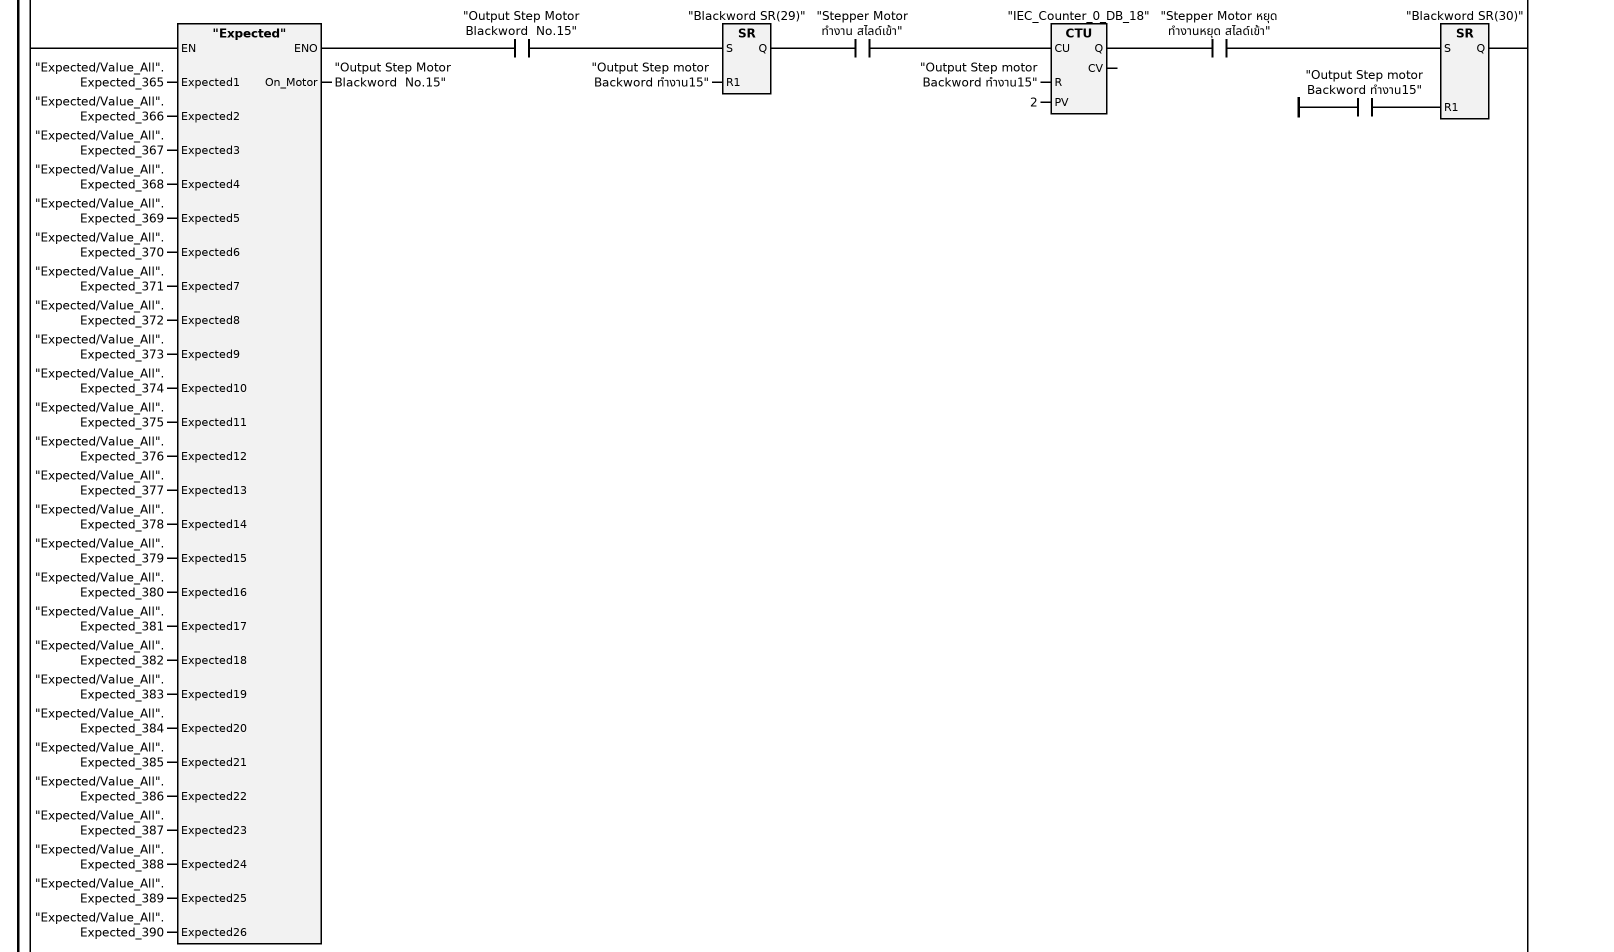
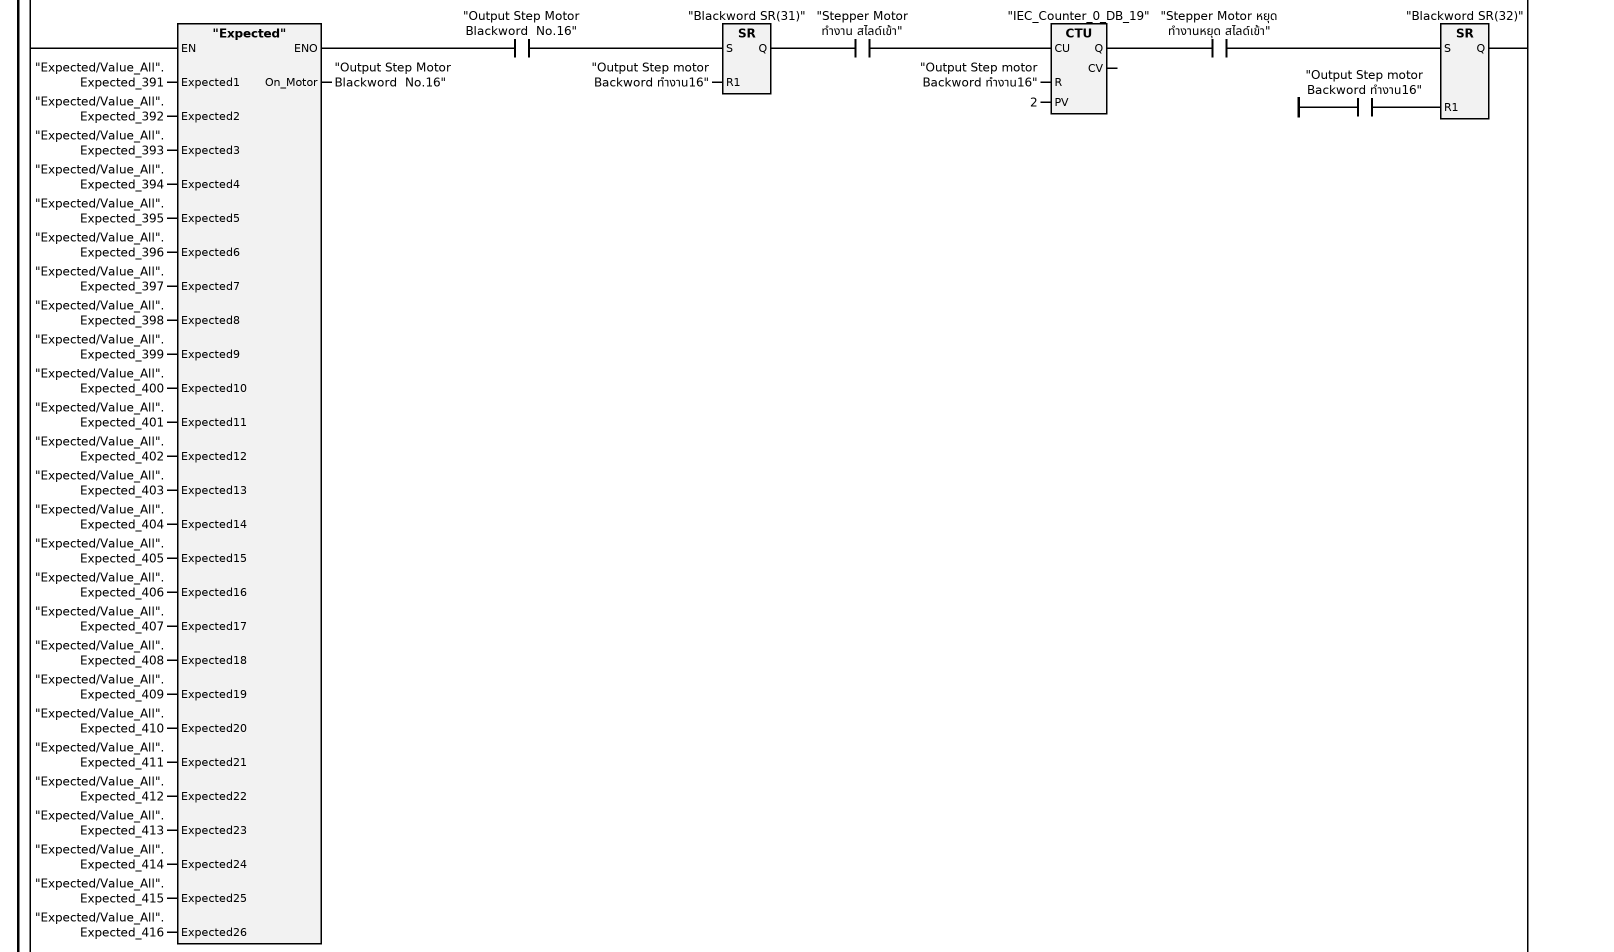
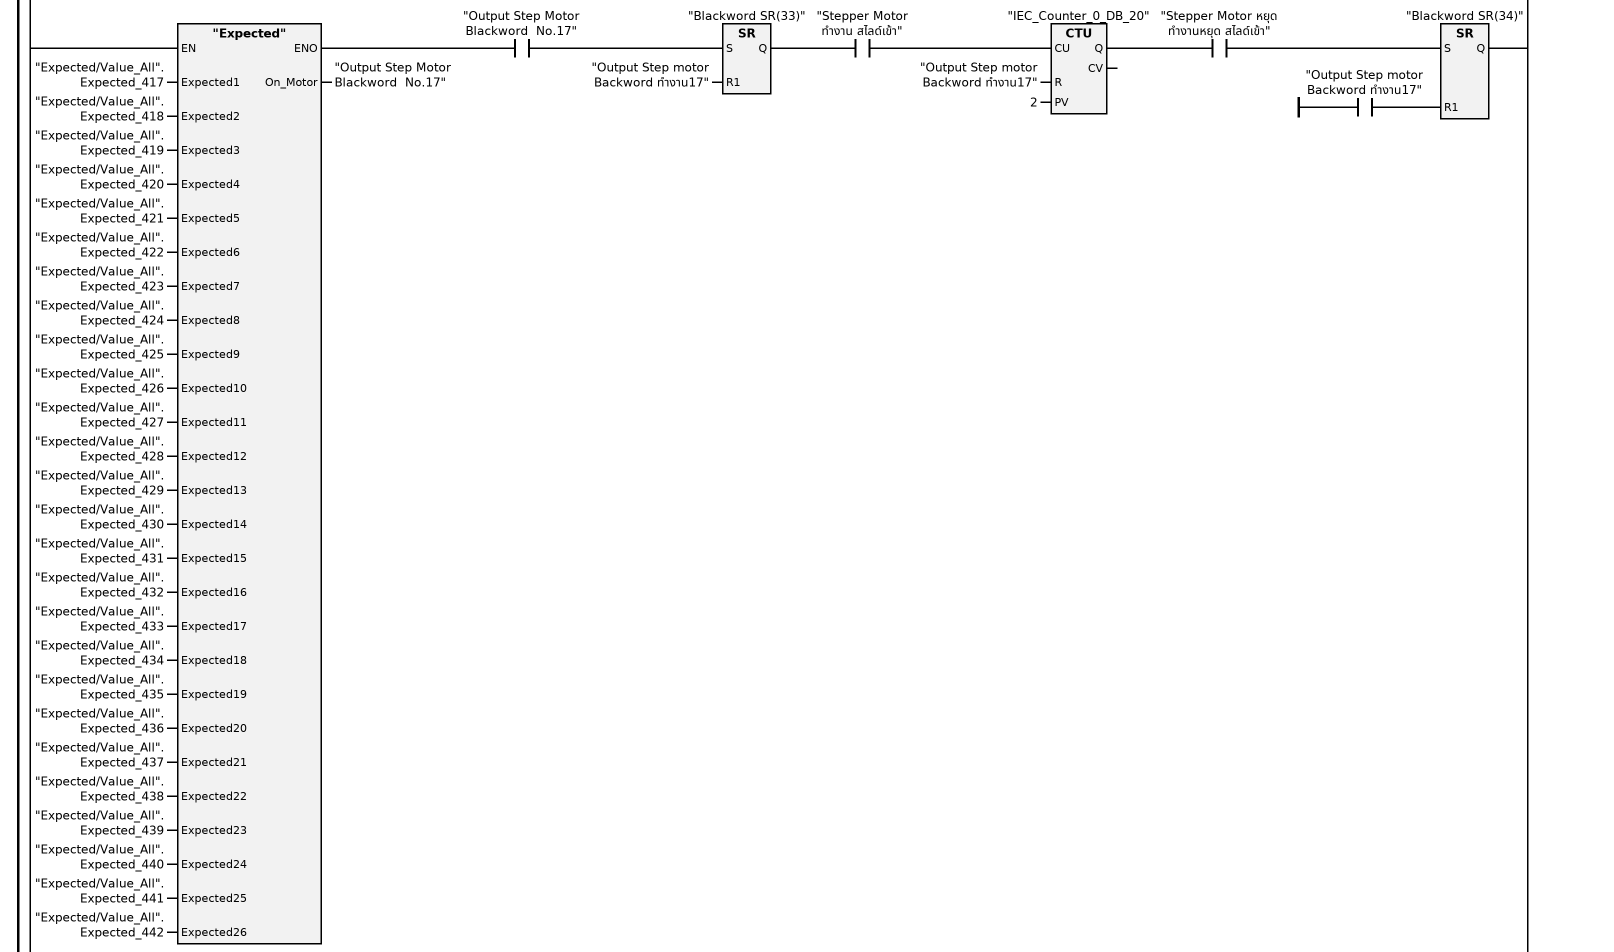
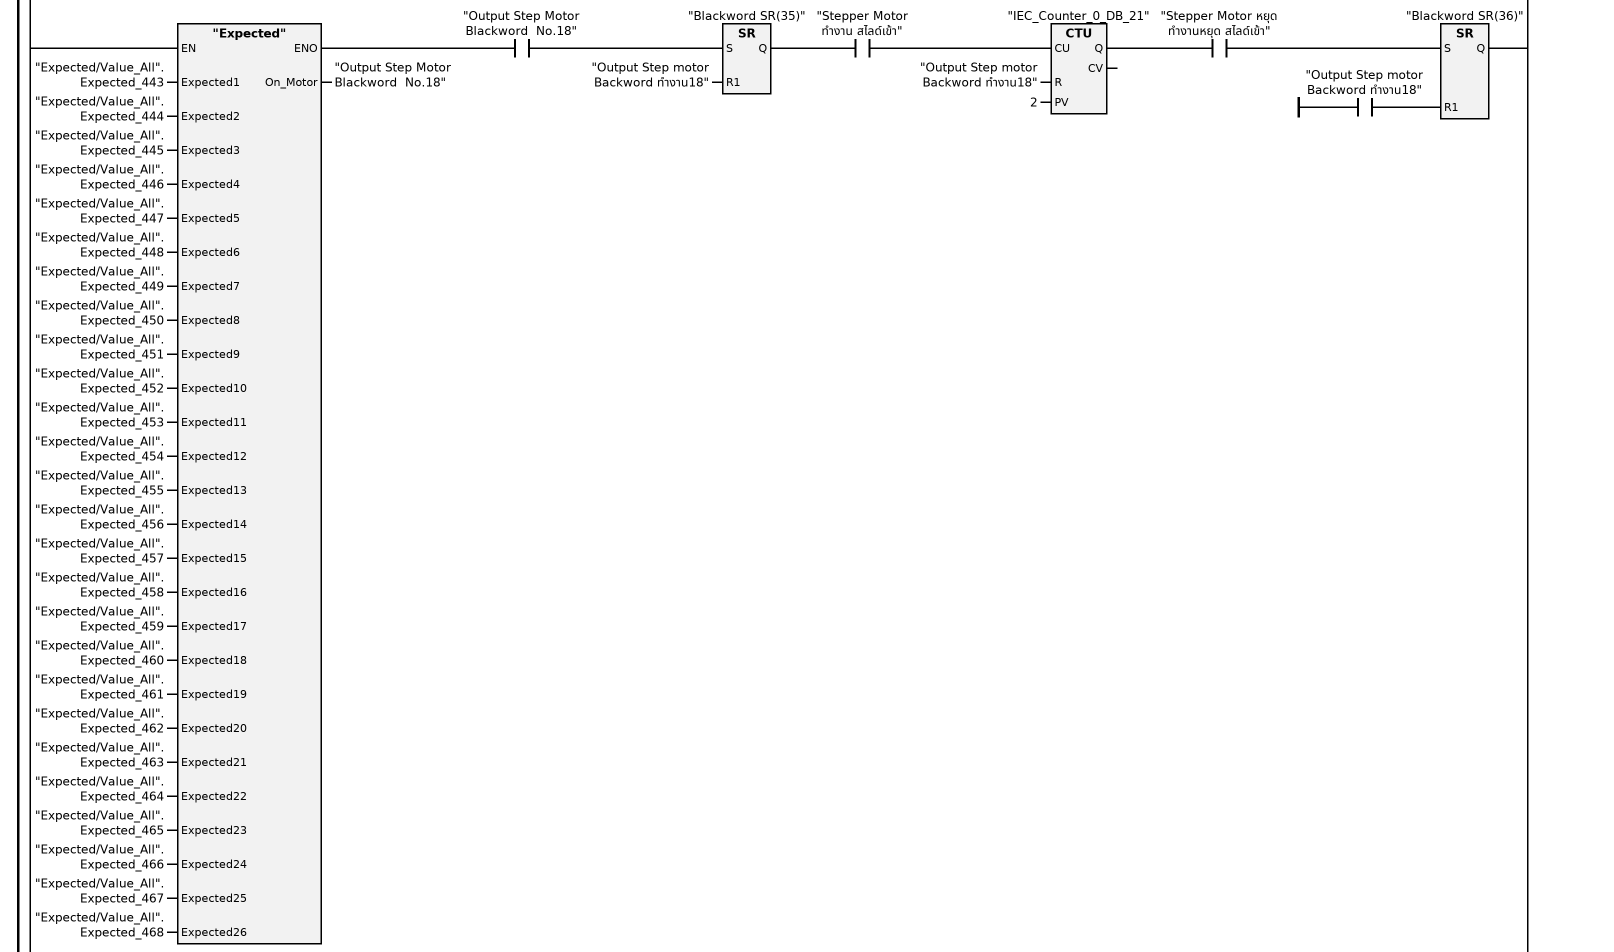
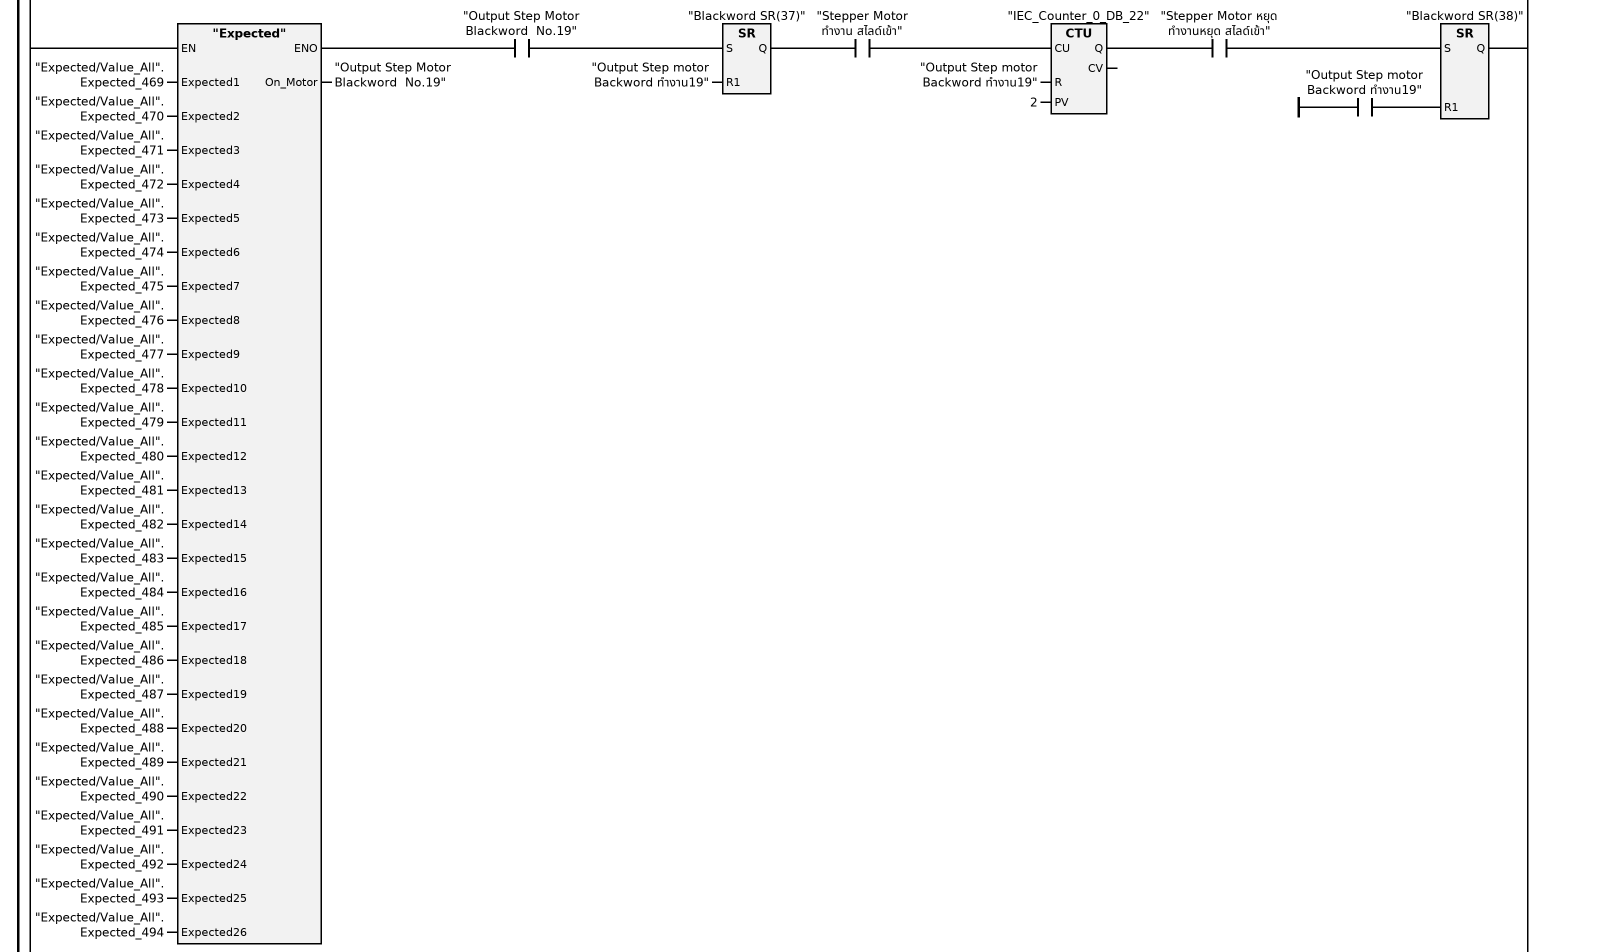
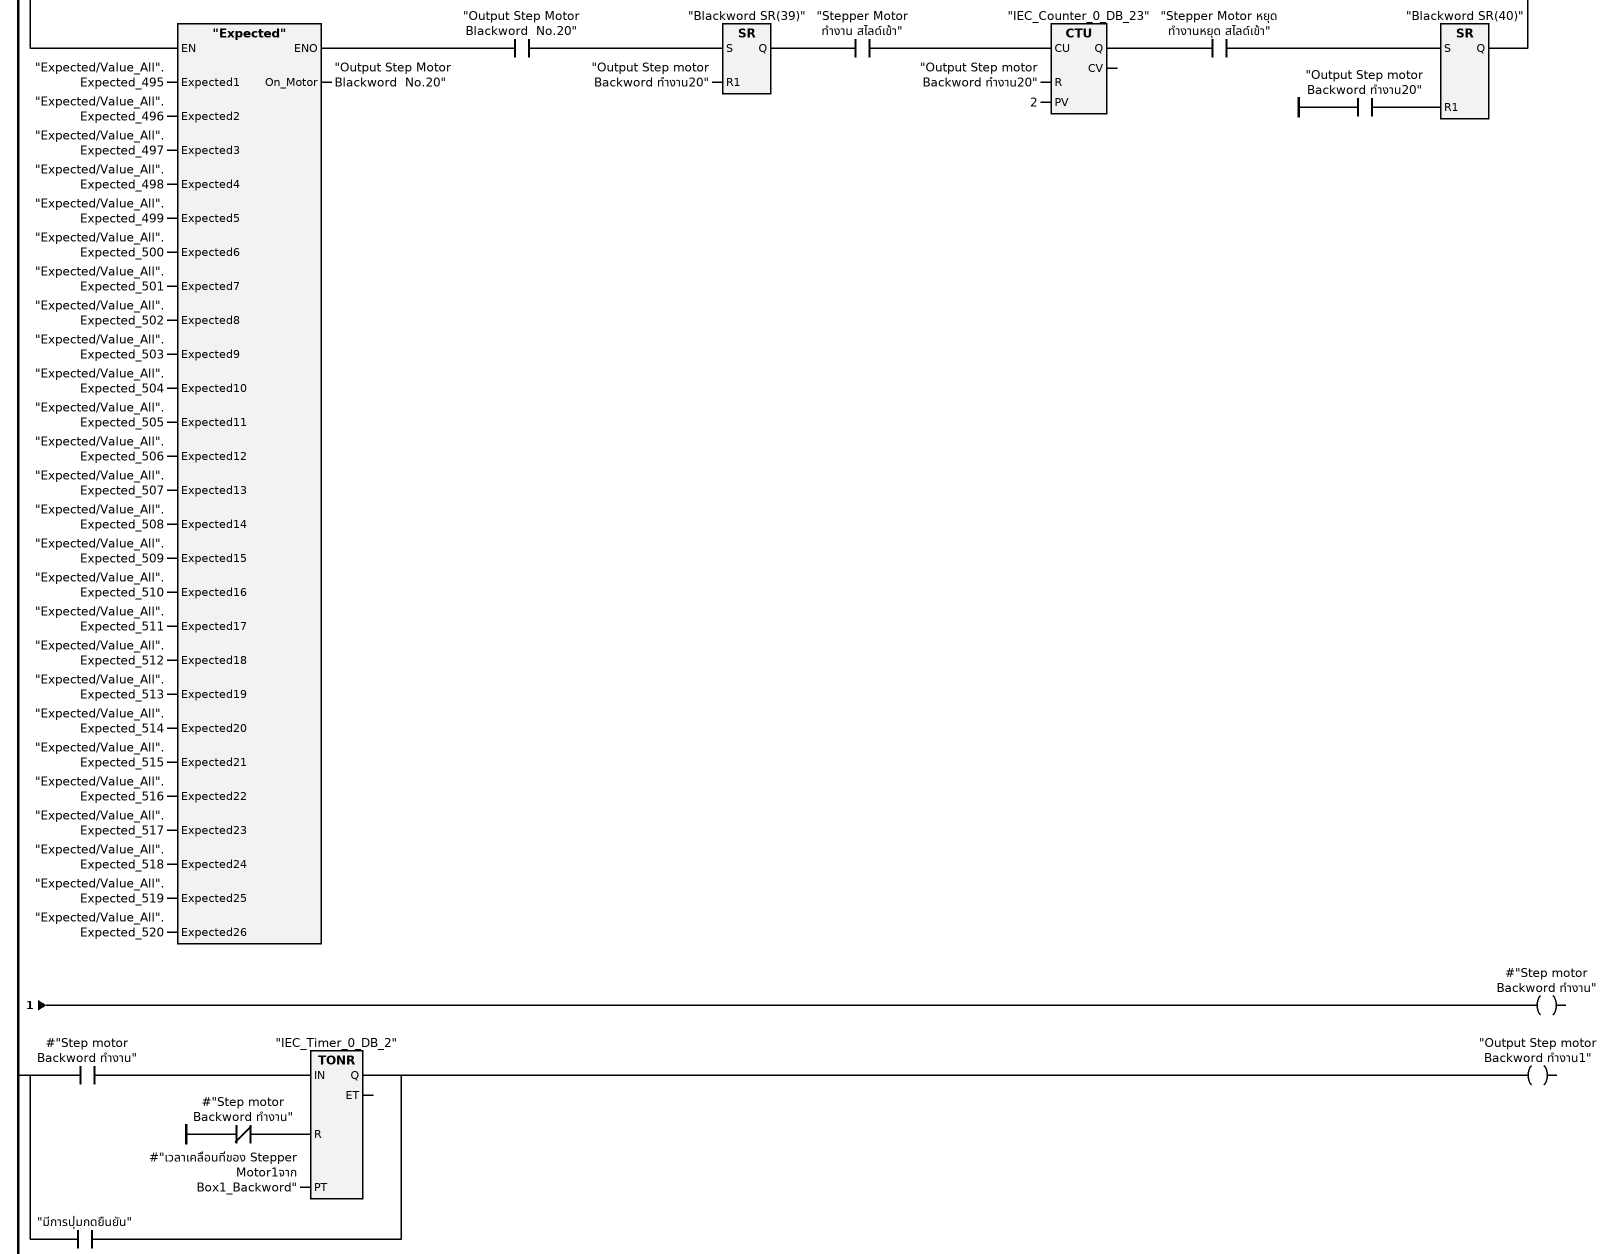
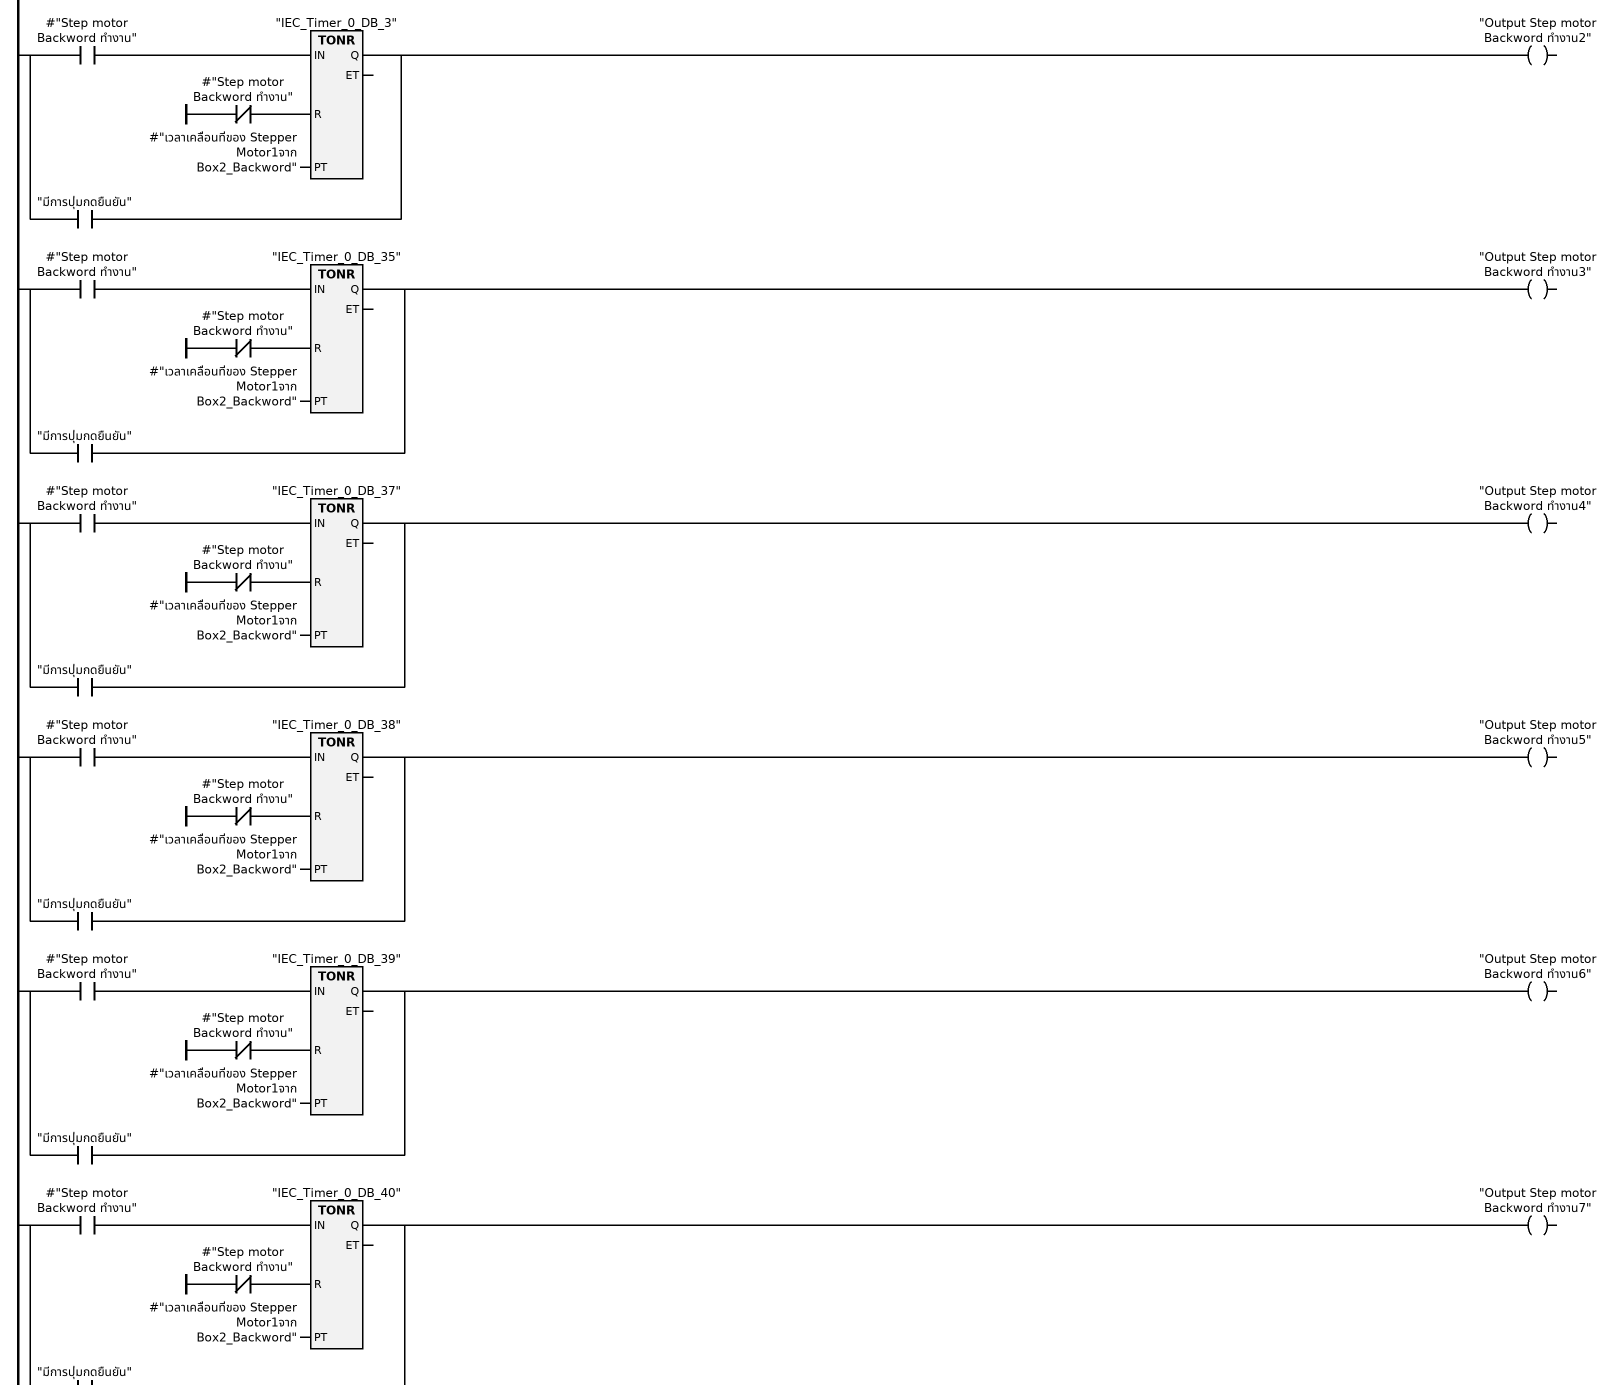
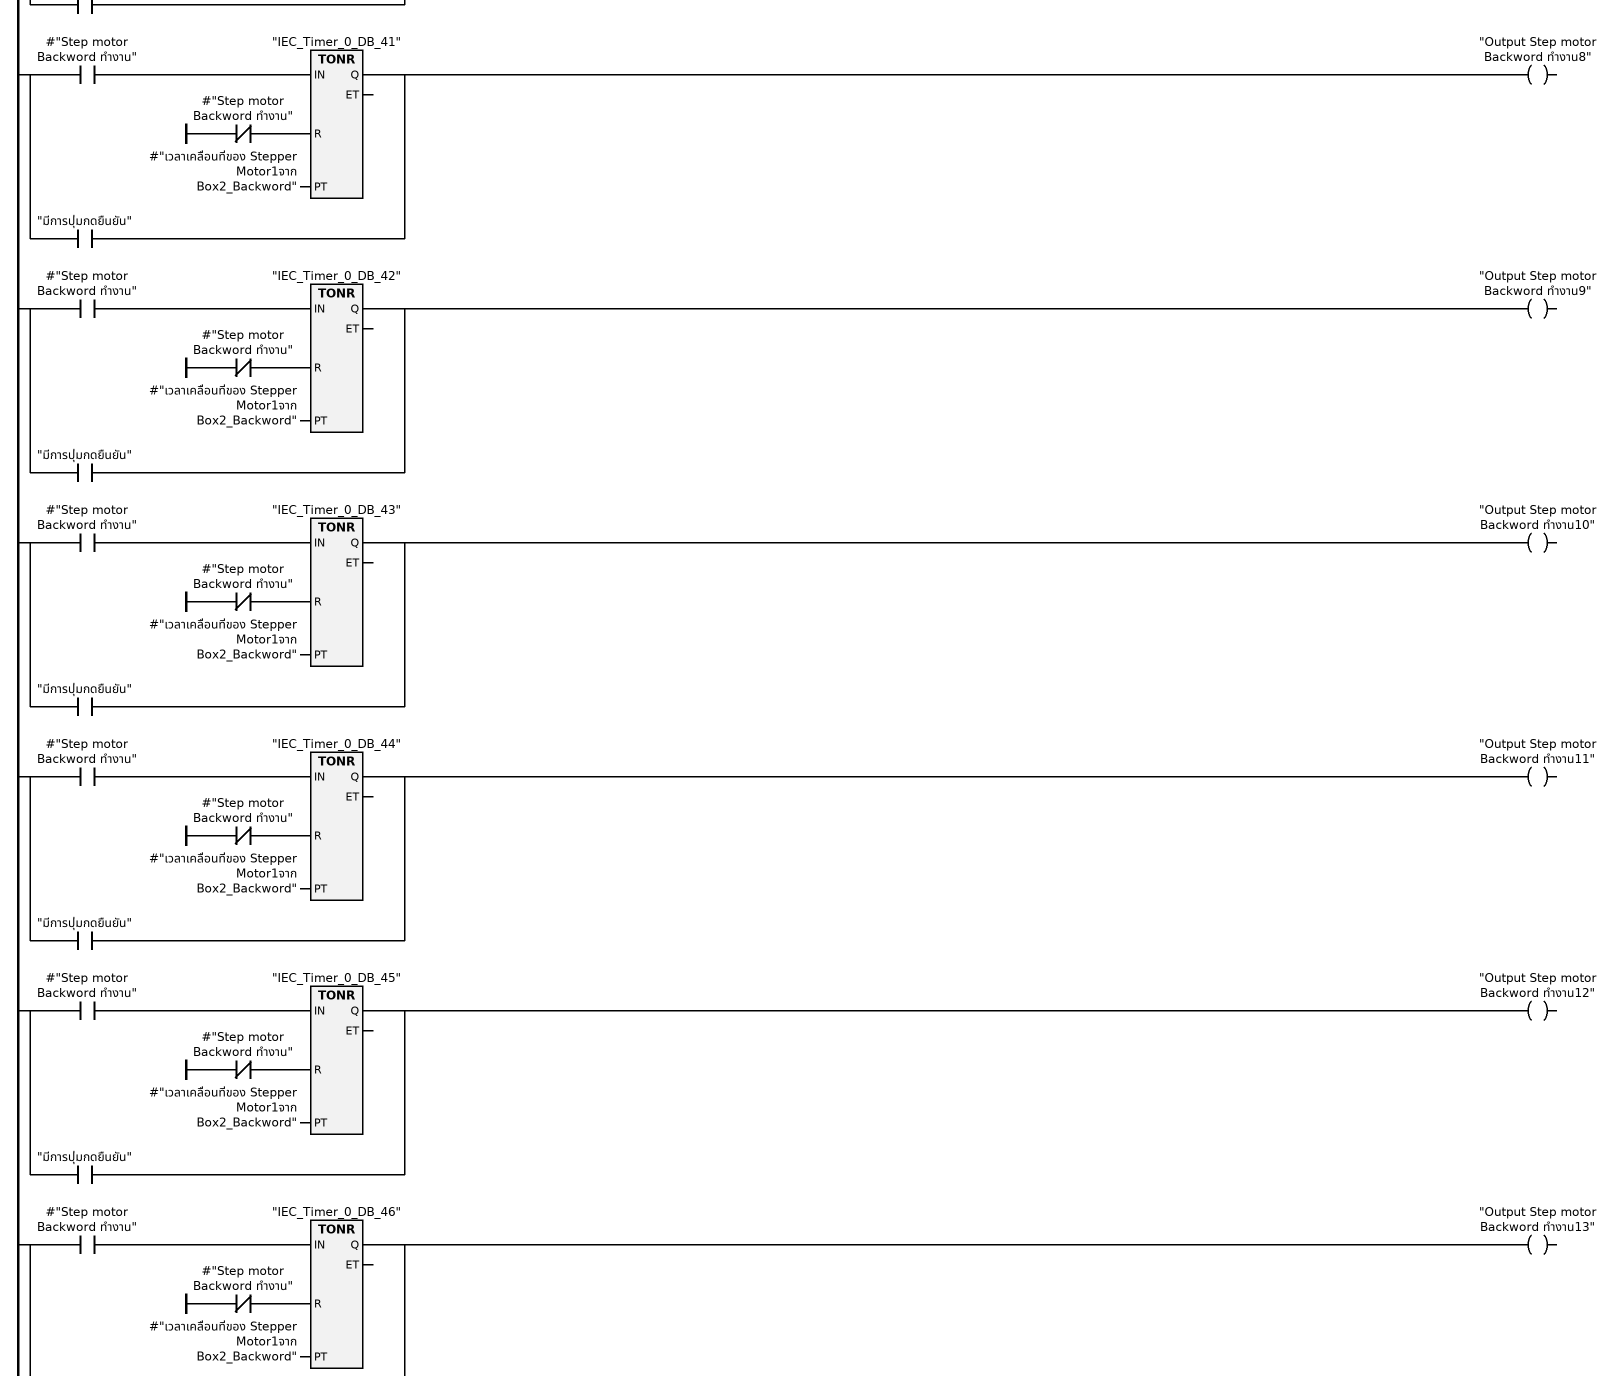
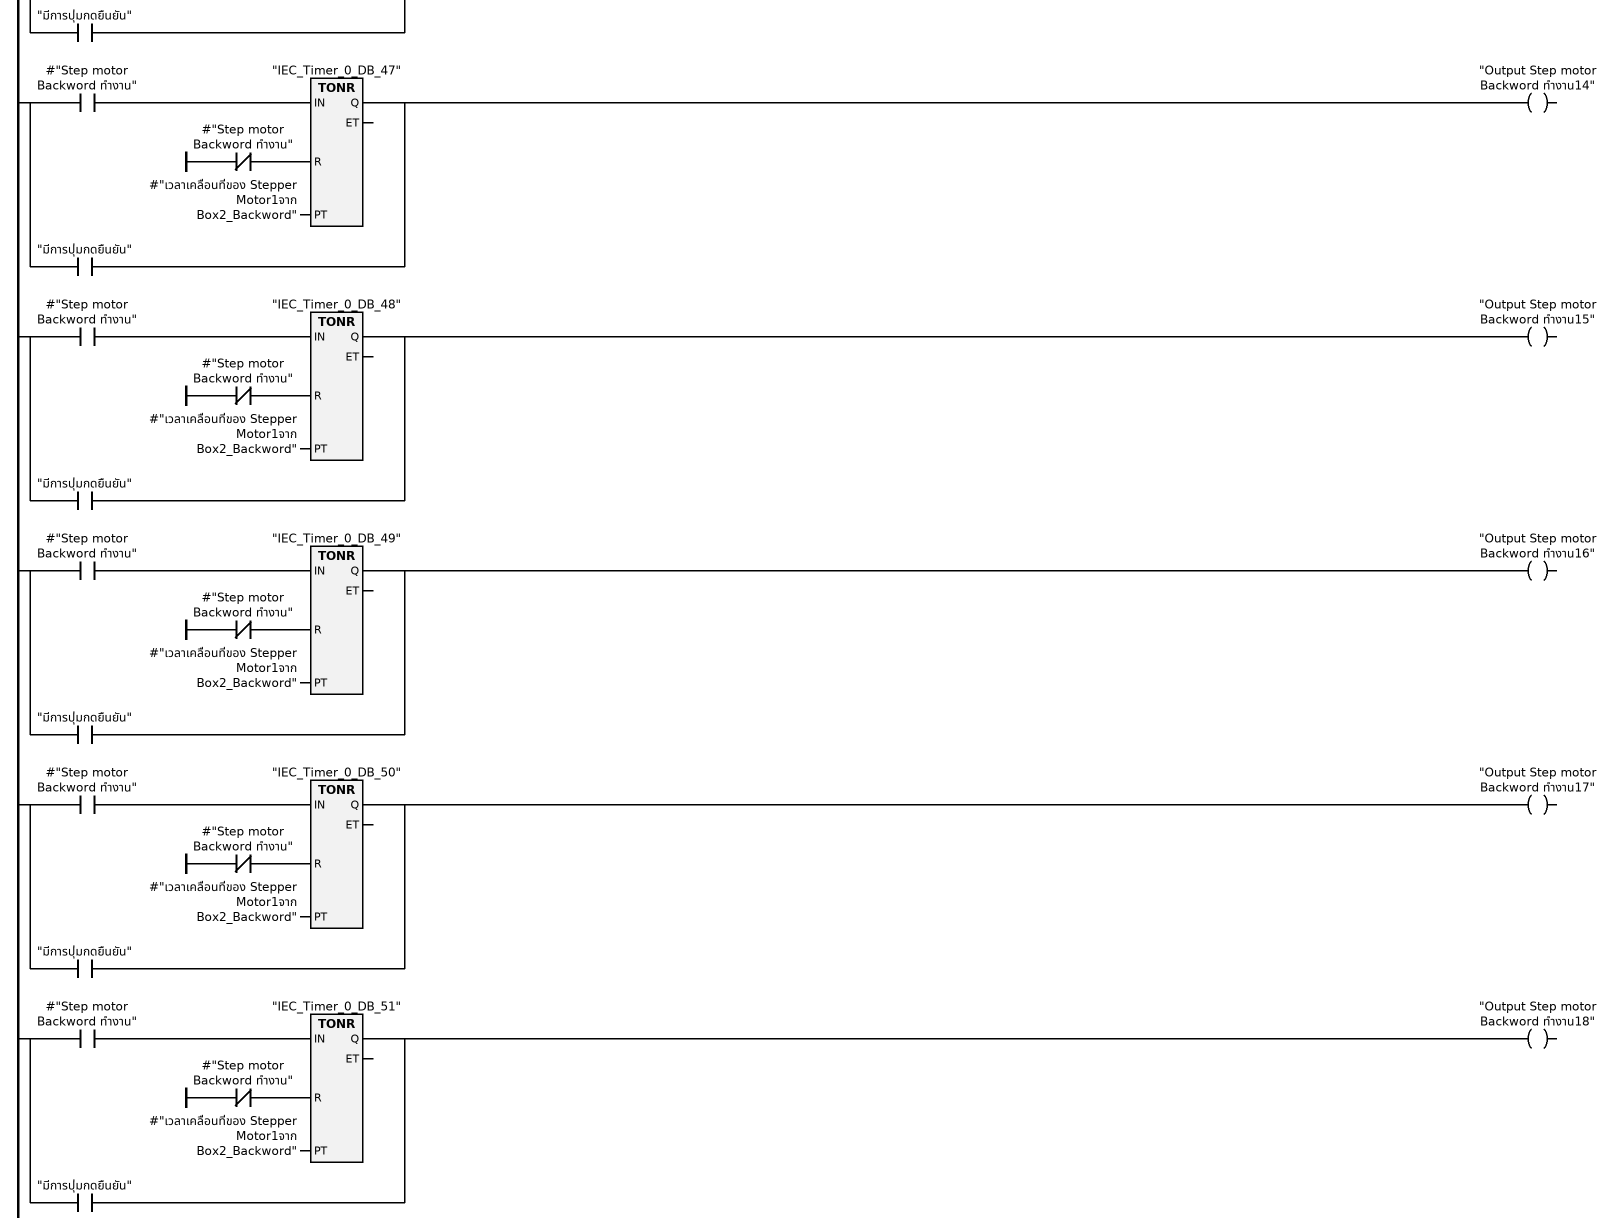
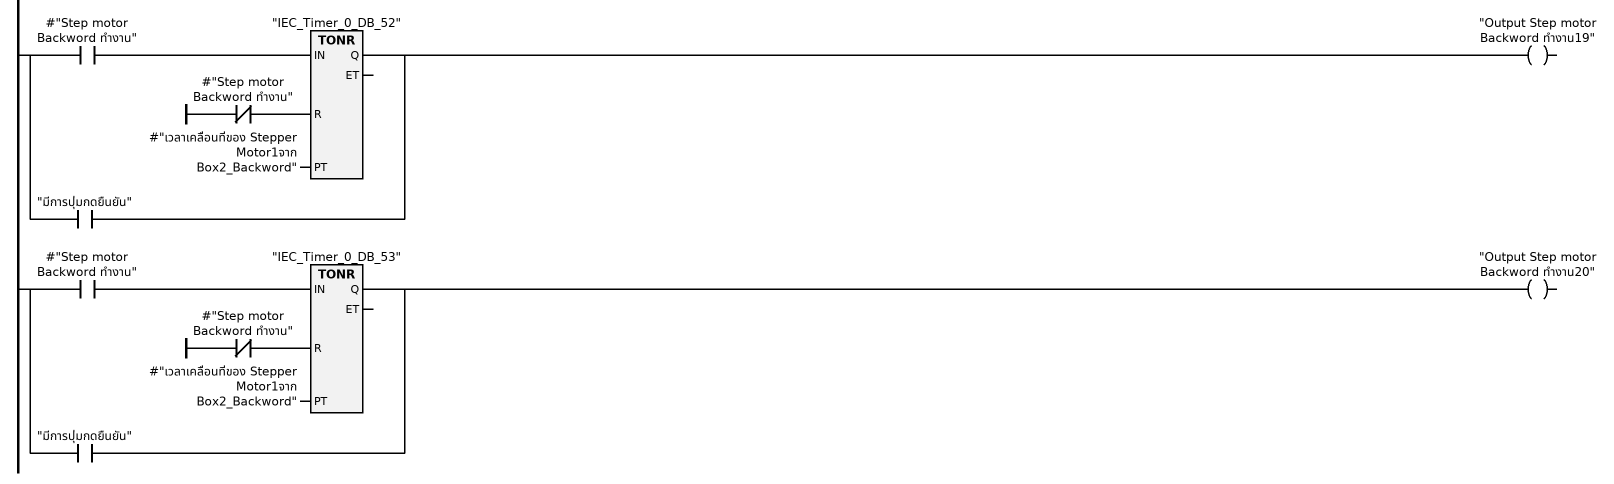
   "Expected"(Expected1 := "Expected/Value_All".Expected_1,
              Expected2 := "Expected/Value_All".Expected_2,
              Expected3 := "Expected/Value_All".Expected_3,
              Expected4 := "Expected/Value_All".Expected_4,
              Expected5 := "Expected/Value_All".Expected_5,
              Expected6 := "Expected/Value_All".Expected_6,
              Expected7 := "Expected/Value_All".Expected_7,
              Expected8 := "Expected/Value_All".Expected_8,
              Expected9 := "Expected/Value_All".Expected_9,
              Expected10 := "Expected/Value_All".Expected_10,
              Expected11 := "Expected/Value_All".Expected_11,
              Expected12 := "Expected/Value_All".Expected_12,
              Expected13 := "Expected/Value_All".Expected_13,
              Expected14 := "Expected/Value_All".Expected_14,
              Expected15 := "Expected/Value_All".Expected_15,
              Expected16 := "Expected/Value_All".Expected_16,
              Expected17 := "Expected/Value_All".Expected_17,
              Expected18 := "Expected/Value_All".Expected_18,
              Expected19 := "Expected/Value_All".Expected_19,
              Expected20 := "Expected/Value_All".Expected_20,
              Expected21 := "Expected/Value_All".Expected_21,
              Expected22 := "Expected/Value_All".Expected_22,
              Expected23 := "Expected/Value_All".Expected_23,
              Expected24 := "Expected/Value_All".Expected_24,
              Expected25 := "Expected/Value_All".Expected_25,
              Expected26 := "Expected/Value_All".Expected_26,
              On_Motor => "Output Step Motor Blackword  No.1",
              ENO => #_w1);
   IF #_w1 AND "Output Step Motor Blackword  No.1" THEN
       "Blackword SR(1)" := TRUE;   // SR flip-flop
   END_IF;
   IF "Output Step motor  Backword ทำงาน1" THEN "Blackword SR(1)" := FALSE; END_IF;
   "IEC_Counter_0_DB_24".CTU(CU := "Blackword SR(1)" AND "Stepper Motor ทำงาน สไลด์เข้า",
                           R := "Output Step motor  Backword ทำงาน1",
                           PV := 2);
   IF "IEC_Counter_0_DB_24".Q AND "Stepper Motor หยุด ทำงานหยุด สไลด์เข้า" THEN
       "Blackword SR(2)" := TRUE;   // SR flip-flop
   END_IF;
   IF "Output Step motor  Backword ทำงาน1" THEN "Blackword SR(2)" := FALSE; END_IF;
   #_w3 := "Blackword SR(2)";
   "Expected"(Expected1 := "Expected/Value_All".Expected_27,
              Expected2 := "Expected/Value_All".Expected_28,
              Expected3 := "Expected/Value_All".Expected_29,
              Expected4 := "Expected/Value_All".Expected_30,
              Expected5 := "Expected/Value_All".Expected_31,
              Expected6 := "Expected/Value_All".Expected_32,
              Expected7 := "Expected/Value_All".Expected_33,
              Expected8 := "Expected/Value_All".Expected_34,
              Expected9 := "Expected/Value_All".Expected_35,
              Expected10 := "Expected/Value_All".Expected_36,
              Expected11 := "Expected/Value_All".Expected_37,
              Expected12 := "Expected/Value_All".Expected_38,
              Expected13 := "Expected/Value_All".Expected_39,
              Expected14 := "Expected/Value_All".Expected_40,
              Expected15 := "Expected/Value_All".Expected_41,
              Expected16 := "Expected/Value_All".Expected_42,
              Expected17 := "Expected/Value_All".Expected_43,
              Expected18 := "Expected/Value_All".Expected_44,
              Expected19 := "Expected/Value_All".Expected_45,
              Expected20 := "Expected/Value_All".Expected_46,
              Expected21 := "Expected/Value_All".Expected_47,
              Expected22 := "Expected/Value_All".Expected_48,
              Expected23 := "Expected/Value_All".Expected_49,
              Expected24 := "Expected/Value_All".Expected_50,
              Expected25 := "Expected/Value_All".Expected_51,
              Expected26 := "Expected/Value_All".Expected_52,
              On_Motor => "Output Step Motor Blackword  No.2",
              ENO => #_w2);
   IF #_w2 AND "Output Step Motor Blackword  No.2" THEN
       "Blackword SR(3)" := TRUE;   // SR flip-flop
   END_IF;
   IF "Output Step motor  Backword ทำงาน2" THEN "Blackword SR(3)" := FALSE; END_IF;
   "IEC_Counter_0_DB_3".CTU(CU := "Blackword SR(3)" AND "Stepper Motor ทำงาน สไลด์เข้า",
                           R := "Output Step motor  Backword ทำงาน2",
                           PV := 2);
   IF "IEC_Counter_0_DB_3".Q AND "Stepper Motor หยุด ทำงานหยุด สไลด์เข้า" THEN
       "Blackword SR(4)" := TRUE;   // SR flip-flop
   END_IF;
   IF "Output Step motor  Backword ทำงาน2" THEN "Blackword SR(4)" := FALSE; END_IF;
   #_w5 := "Blackword SR(4)";
   "Expected"(Expected1 := "Expected/Value_All".Expected_53,
              Expected2 := "Expected/Value_All".Expected_54,
              Expected3 := "Expected/Value_All".Expected_55,
              Expected4 := "Expected/Value_All".Expected_56,
              Expected5 := "Expected/Value_All".Expected_57,
              Expected6 := "Expected/Value_All".Expected_58,
              Expected7 := "Expected/Value_All".Expected_59,
              Expected8 := "Expected/Value_All".Expected_60,
              Expected9 := "Expected/Value_All".Expected_61,
              Expected10 := "Expected/Value_All".Expected_62,
              Expected11 := "Expected/Value_All".Expected_63,
              Expected12 := "Expected/Value_All".Expected_64,
              Expected13 := "Expected/Value_All".Expected_65,
              Expected14 := "Expected/Value_All".Expected_66,
              Expected15 := "Expected/Value_All".Expected_67,
              Expected16 := "Expected/Value_All".Expected_68,
              Expected17 := "Expected/Value_All".Expected_69,
              Expected18 := "Expected/Value_All".Expected_70,
              Expected19 := "Expected/Value_All".Expected_71,
              Expected20 := "Expected/Value_All".Expected_72,
              Expected21 := "Expected/Value_All".Expected_73,
              Expected22 := "Expected/Value_All".Expected_74,
              Expected23 := "Expected/Value_All".Expected_75,
              Expected24 := "Expected/Value_All".Expected_76,
              Expected25 := "Expected/Value_All".Expected_77,
              Expected26 := "Expected/Value_All".Expected_78,
              On_Motor => "Output Step Motor Blackword  No.3",
              ENO => #_w4);
   IF #_w4 AND "Output Step Motor Blackword  No.3" THEN
       "Blackword SR(5)" := TRUE;   // SR flip-flop
   END_IF;
   IF "Output Step motor  Backword ทำงาน3" THEN "Blackword SR(5)" := FALSE; END_IF;
   "IEC_Counter_0_DB_4".CTU(CU := "Blackword SR(5)" AND "Stepper Motor ทำงาน สไลด์เข้า",
                           R := "Output Step motor  Backword ทำงาน3",
                           PV := 2);
   IF "IEC_Counter_0_DB_4".Q AND "Stepper Motor หยุด ทำงานหยุด สไลด์เข้า" THEN
       "Blackword SR(6)" := TRUE;   // SR flip-flop
   END_IF;
   IF "Output Step motor  Backword ทำงาน3" THEN "Blackword SR(6)" := FALSE; END_IF;
   #_w7 := "Blackword SR(6)";
   "Expected"(Expected1 := "Expected/Value_All".Expected_79,
              Expected2 := "Expected/Value_All".Expected_80,
              Expected3 := "Expected/Value_All".Expected_81,
              Expected4 := "Expected/Value_All".Expected_82,
              Expected5 := "Expected/Value_All".Expected_83,
              Expected6 := "Expected/Value_All".Expected_84,
              Expected7 := "Expected/Value_All".Expected_85,
              Expected8 := "Expected/Value_All".Expected_86,
              Expected9 := "Expected/Value_All".Expected_87,
              Expected10 := "Expected/Value_All".Expected_88,
              Expected11 := "Expected/Value_All".Expected_89,
              Expected12 := "Expected/Value_All".Expected_90,
              Expected13 := "Expected/Value_All".Expected_91,
              Expected14 := "Expected/Value_All".Expected_92,
              Expected15 := "Expected/Value_All".Expected_93,
              Expected16 := "Expected/Value_All".Expected_94,
              Expected17 := "Expected/Value_All".Expected_95,
              Expected18 := "Expected/Value_All".Expected_96,
              Expected19 := "Expected/Value_All".Expected_97,
              Expected20 := "Expected/Value_All".Expected_98,
              Expected21 := "Expected/Value_All".Expected_99,
              Expected22 := "Expected/Value_All".Expected_100,
              Expected23 := "Expected/Value_All".Expected_101,
              Expected24 := "Expected/Value_All".Expected_102,
              Expected25 := "Expected/Value_All".Expected_103,
              Expected26 := "Expected/Value_All".Expected_104,
              On_Motor => "Output Step Motor Blackword  No.4",
              ENO => #_w6);
   IF #_w6 AND "Output Step Motor Blackword  No.4" THEN
       "Blackword SR(7)" := TRUE;   // SR flip-flop
   END_IF;
   IF "Output Step motor  Backword ทำงาน4" THEN "Blackword SR(7)" := FALSE; END_IF;
   "IEC_Counter_0_DB_7".CTU(CU := "Blackword SR(7)" AND "Stepper Motor ทำงาน สไลด์เข้า",
                           R := "Output Step motor  Backword ทำงาน4",
                           PV := 2);
   IF "IEC_Counter_0_DB_7".Q AND "Stepper Motor หยุด ทำงานหยุด สไลด์เข้า" THEN
       "Blackword SR(8)" := TRUE;   // SR flip-flop
   END_IF;
   IF "Output Step motor  Backword ทำงาน4" THEN "Blackword SR(8)" := FALSE; END_IF;
   #_w9 := "Blackword SR(8)";
   "Expected"(Expected1 := "Expected/Value_All".Expected_105,
              Expected2 := "Expected/Value_All".Expected_106,
              Expected3 := "Expected/Value_All".Expected_107,
              Expected4 := "Expected/Value_All".Expected_108,
              Expected5 := "Expected/Value_All".Expected_109,
              Expected6 := "Expected/Value_All".Expected_110,
              Expected7 := "Expected/Value_All".Expected_111,
              Expected8 := "Expected/Value_All".Expected_112,
              Expected9 := "Expected/Value_All".Expected_113,
              Expected10 := "Expected/Value_All".Expected_114,
              Expected11 := "Expected/Value_All".Expected_115,
              Expected12 := "Expected/Value_All".Expected_116,
              Expected13 := "Expected/Value_All".Expected_117,
              Expected14 := "Expected/Value_All".Expected_118,
              Expected15 := "Expected/Value_All".Expected_119,
              Expected16 := "Expected/Value_All".Expected_120,
              Expected17 := "Expected/Value_All".Expected_121,
              Expected18 := "Expected/Value_All".Expected_122,
              Expected19 := "Expected/Value_All".Expected_123,
              Expected20 := "Expected/Value_All".Expected_124,
              Expected21 := "Expected/Value_All".Expected_125,
              Expected22 := "Expected/Value_All".Expected_126,
              Expected23 := "Expected/Value_All".Expected_127,
              Expected24 := "Expected/Value_All".Expected_128,
              Expected25 := "Expected/Value_All".Expected_129,
              Expected26 := "Expected/Value_All".Expected_130,
              On_Motor => "Output Step Motor Blackword  No.5",
              ENO => #_w8);
   IF #_w8 AND "Output Step Motor Blackword  No.5" THEN
       "Blackword SR(9)" := TRUE;   // SR flip-flop
   END_IF;
   IF "Output Step motor  Backword ทำงาน5" THEN "Blackword SR(9)" := FALSE; END_IF;
   "IEC_Counter_0_DB_8".CTU(CU := "Blackword SR(9)" AND "Stepper Motor ทำงาน สไลด์เข้า",
                           R := "Output Step motor  Backword ทำงาน5",
                           PV := 2);
   IF "IEC_Counter_0_DB_8".Q AND "Stepper Motor หยุด ทำงานหยุด สไลด์เข้า" THEN
       "Blackword SR(10)" := TRUE;   // SR flip-flop
   END_IF;
   IF "Output Step motor  Backword ทำงาน5" THEN "Blackword SR(10)" := FALSE; END_IF;
   #_w11 := "Blackword SR(10)";
   "Expected"(Expected1 := "Expected/Value_All".Expected_131,
              Expected2 := "Expected/Value_All".Expected_132,
              Expected3 := "Expected/Value_All".Expected_133,
              Expected4 := "Expected/Value_All".Expected_134,
              Expected5 := "Expected/Value_All".Expected_135,
              Expected6 := "Expected/Value_All".Expected_136,
              Expected7 := "Expected/Value_All".Expected_137,
              Expected8 := "Expected/Value_All".Expected_138,
              Expected9 := "Expected/Value_All".Expected_139,
              Expected10 := "Expected/Value_All".Expected_140,
              Expected11 := "Expected/Value_All".Expected_141,
              Expected12 := "Expected/Value_All".Expected_142,
              Expected13 := "Expected/Value_All".Expected_143,
              Expected14 := "Expected/Value_All".Expected_144,
              Expected15 := "Expected/Value_All".Expected_145,
              Expected16 := "Expected/Value_All".Expected_146,
              Expected17 := "Expected/Value_All".Expected_147,
              Expected18 := "Expected/Value_All".Expected_148,
              Expected19 := "Expected/Value_All".Expected_149,
              Expected20 := "Expected/Value_All".Expected_150,
              Expected21 := "Expected/Value_All".Expected_151,
              Expected22 := "Expected/Value_All".Expected_152,
              Expected23 := "Expected/Value_All".Expected_153,
              Expected24 := "Expected/Value_All".Expected_154,
              Expected25 := "Expected/Value_All".Expected_155,
              Expected26 := "Expected/Value_All".Expected_156,
              On_Motor => "Output Step Motor Blackword  No.6",
              ENO => #_w10);
   IF #_w10 AND "Output Step Motor Blackword  No.6" THEN
       "Blackword SR(11)" := TRUE;   // SR flip-flop
   END_IF;
   IF "Output Step motor  Backword ทำงาน6" THEN "Blackword SR(11)" := FALSE; END_IF;
   "IEC_Counter_0_DB_9".CTU(CU := "Blackword SR(11)" AND "Stepper Motor ทำงาน สไลด์เข้า",
                           R := "Output Step motor  Backword ทำงาน6",
                           PV := 2);
   IF "IEC_Counter_0_DB_9".Q AND "Stepper Motor หยุด ทำงานหยุด สไลด์เข้า" THEN
       "Blackword SR(12)" := TRUE;   // SR flip-flop
   END_IF;
   IF "Output Step motor  Backword ทำงาน6" THEN "Blackword SR(12)" := FALSE; END_IF;
   #_w13 := "Blackword SR(12)";
   "Expected"(Expected1 := "Expected/Value_All".Expected_157,
              Expected2 := "Expected/Value_All".Expected_158,
              Expected3 := "Expected/Value_All".Expected_159,
              Expected4 := "Expected/Value_All".Expected_160,
              Expected5 := "Expected/Value_All".Expected_161,
              Expected6 := "Expected/Value_All".Expected_162,
              Expected7 := "Expected/Value_All".Expected_163,
              Expected8 := "Expected/Value_All".Expected_164,
              Expected9 := "Expected/Value_All".Expected_165,
              Expected10 := "Expected/Value_All".Expected_166,
              Expected11 := "Expected/Value_All".Expected_167,
              Expected12 := "Expected/Value_All".Expected_168,
              Expected13 := "Expected/Value_All".Expected_169,
              Expected14 := "Expected/Value_All".Expected_170,
              Expected15 := "Expected/Value_All".Expected_171,
              Expected16 := "Expected/Value_All".Expected_172,
              Expected17 := "Expected/Value_All".Expected_173,
              Expected18 := "Expected/Value_All".Expected_174,
              Expected19 := "Expected/Value_All".Expected_175,
              Expected20 := "Expected/Value_All".Expected_176,
              Expected21 := "Expected/Value_All".Expected_177,
              Expected22 := "Expected/Value_All".Expected_178,
              Expected23 := "Expected/Value_All".Expected_179,
              Expected24 := "Expected/Value_All".Expected_180,
              Expected25 := "Expected/Value_All".Expected_181,
              Expected26 := "Expected/Value_All".Expected_182,
              On_Motor => "Output Step Motor Blackword  No.7",
              ENO => #_w12);
   IF #_w12 AND "Output Step Motor Blackword  No.7" THEN
       "Blackword SR(13)" := TRUE;   // SR flip-flop
   END_IF;
   IF "Output Step motor  Backword ทำงาน7" THEN "Blackword SR(13)" := FALSE; END_IF;
   "IEC_Counter_0_DB_10".CTU(CU := "Blackword SR(13)" AND "Stepper Motor ทำงาน สไลด์เข้า",
                           R := "Output Step motor  Backword ทำงาน7",
                           PV := 2);
   IF "IEC_Counter_0_DB_10".Q AND "Stepper Motor หยุด ทำงานหยุด สไลด์เข้า" THEN
       "Blackword SR(14)" := TRUE;   // SR flip-flop
   END_IF;
   IF "Output Step motor  Backword ทำงาน7" THEN "Blackword SR(14)" := FALSE; END_IF;
   #_w15 := "Blackword SR(14)";
   "Expected"(Expected1 := "Expected/Value_All".Expected_183,
              Expected2 := "Expected/Value_All".Expected_184,
              Expected3 := "Expected/Value_All".Expected_185,
              Expected4 := "Expected/Value_All".Expected_186,
              Expected5 := "Expected/Value_All".Expected_187,
              Expected6 := "Expected/Value_All".Expected_188,
              Expected7 := "Expected/Value_All".Expected_189,
              Expected8 := "Expected/Value_All".Expected_190,
              Expected9 := "Expected/Value_All".Expected_191,
              Expected10 := "Expected/Value_All".Expected_192,
              Expected11 := "Expected/Value_All".Expected_193,
              Expected12 := "Expected/Value_All".Expected_194,
              Expected13 := "Expected/Value_All".Expected_195,
              Expected14 := "Expected/Value_All".Expected_196,
              Expected15 := "Expected/Value_All".Expected_197,
              Expected16 := "Expected/Value_All".Expected_198,
              Expected17 := "Expected/Value_All".Expected_199,
              Expected18 := "Expected/Value_All".Expected_200,
              Expected19 := "Expected/Value_All".Expected_201,
              Expected20 := "Expected/Value_All".Expected_202,
              Expected21 := "Expected/Value_All".Expected_203,
              Expected22 := "Expected/Value_All".Expected_204,
              Expected23 := "Expected/Value_All".Expected_205,
              Expected24 := "Expected/Value_All".Expected_206,
              Expected25 := "Expected/Value_All".Expected_207,
              Expected26 := "Expected/Value_All".Expected_208,
              On_Motor => "Output Step Motor Blackword  No.8",
              ENO => #_w14);
   IF #_w14 AND "Output Step Motor Blackword  No.8" THEN
       "Blackword SR(15)" := TRUE;   // SR flip-flop
   END_IF;
   IF "Output Step motor  Backword ทำงาน8" THEN "Blackword SR(15)" := FALSE; END_IF;
   "IEC_Counter_0_DB_11".CTU(CU := "Blackword SR(15)" AND "Stepper Motor ทำงาน สไลด์เข้า",
                           R := "Output Step motor  Backword ทำงาน8",
                           PV := 2);
   IF "IEC_Counter_0_DB_11".Q AND "Stepper Motor หยุด ทำงานหยุด สไลด์เข้า" THEN
       "Blackword SR(16)" := TRUE;   // SR flip-flop
   END_IF;
   IF "Output Step motor  Backword ทำงาน8" THEN "Blackword SR(16)" := FALSE; END_IF;
   #_w17 := "Blackword SR(16)";
   "Expected"(Expected1 := "Expected/Value_All".Expected_209,
              Expected2 := "Expected/Value_All".Expected_210,
              Expected3 := "Expected/Value_All".Expected_211,
              Expected4 := "Expected/Value_All".Expected_212,
              Expected5 := "Expected/Value_All".Expected_213,
              Expected6 := "Expected/Value_All".Expected_214,
              Expected7 := "Expected/Value_All".Expected_215,
              Expected8 := "Expected/Value_All".Expected_216,
              Expected9 := "Expected/Value_All".Expected_217,
              Expected10 := "Expected/Value_All".Expected_218,
              Expected11 := "Expected/Value_All".Expected_219,
              Expected12 := "Expected/Value_All".Expected_220,
              Expected13 := "Expected/Value_All".Expected_221,
              Expected14 := "Expected/Value_All".Expected_222,
              Expected15 := "Expected/Value_All".Expected_223,
              Expected16 := "Expected/Value_All".Expected_224,
              Expected17 := "Expected/Value_All".Expected_225,
              Expected18 := "Expected/Value_All".Expected_226,
              Expected19 := "Expected/Value_All".Expected_227,
              Expected20 := "Expected/Value_All".Expected_228,
              Expected21 := "Expected/Value_All".Expected_229,
              Expected22 := "Expected/Value_All".Expected_230,
              Expected23 := "Expected/Value_All".Expected_231,
              Expected24 := "Expected/Value_All".Expected_232,
              Expected25 := "Expected/Value_All".Expected_233,
              Expected26 := "Expected/Value_All".Expected_234,
              On_Motor => "Output Step Motor Blackword  No.9",
              ENO => #_w16);
   IF #_w16 AND "Output Step Motor Blackword  No.9" THEN
       "Blackword SR(17)" := TRUE;   // SR flip-flop
   END_IF;
   IF "Output Step motor  Backword ทำงาน9" THEN "Blackword SR(17)" := FALSE; END_IF;
   "IEC_Counter_0_DB_12".CTU(CU := "Blackword SR(17)" AND "Stepper Motor ทำงาน สไลด์เข้า",
                           R := "Output Step motor  Backword ทำงาน9",
                           PV := 2);
   IF "IEC_Counter_0_DB_12".Q AND "Stepper Motor หยุด ทำงานหยุด สไลด์เข้า" THEN
       "Blackword SR(18)" := TRUE;   // SR flip-flop
   END_IF;
   IF "Output Step motor  Backword ทำงาน9" THEN "Blackword SR(18)" := FALSE; END_IF;
   #_w19 := "Blackword SR(18)";
   "Expected"(Expected1 := "Expected/Value_All".Expected_235,
              Expected2 := "Expected/Value_All".Expected_236,
              Expected3 := "Expected/Value_All".Expected_237,
              Expected4 := "Expected/Value_All".Expected_238,
              Expected5 := "Expected/Value_All".Expected_239,
              Expected6 := "Expected/Value_All".Expected_240,
              Expected7 := "Expected/Value_All".Expected_241,
              Expected8 := "Expected/Value_All".Expected_242,
              Expected9 := "Expected/Value_All".Expected_243,
              Expected10 := "Expected/Value_All".Expected_244,
              Expected11 := "Expected/Value_All".Expected_245,
              Expected12 := "Expected/Value_All".Expected_246,
              Expected13 := "Expected/Value_All".Expected_247,
              Expected14 := "Expected/Value_All".Expected_248,
              Expected15 := "Expected/Value_All".Expected_249,
              Expected16 := "Expected/Value_All".Expected_250,
              Expected17 := "Expected/Value_All".Expected_251,
              Expected18 := "Expected/Value_All".Expected_252,
              Expected19 := "Expected/Value_All".Expected_253,
              Expected20 := "Expected/Value_All".Expected_254,
              Expected21 := "Expected/Value_All".Expected_255,
              Expected22 := "Expected/Value_All".Expected_256,
              Expected23 := "Expected/Value_All".Expected_257,
              Expected24 := "Expected/Value_All".Expected_258,
              Expected25 := "Expected/Value_All".Expected_259,
              Expected26 := "Expected/Value_All".Expected_260,
              On_Motor => "Output Step Motor Blackword  No.10",
              ENO => #_w18);
   IF #_w18 AND "Output Step Motor Blackword  No.10" THEN
       "Blackword SR(19)" := TRUE;   // SR flip-flop
   END_IF;
   IF "Output Step motor  Backword ทำงาน10" THEN "Blackword SR(19)" := FALSE; END_IF;
   "IEC_Counter_0_DB_13".CTU(CU := "Blackword SR(19)" AND "Stepper Motor ทำงาน สไลด์เข้า",
                           R := "Output Step motor  Backword ทำงาน10",
                           PV := 2);
   IF "IEC_Counter_0_DB_13".Q AND "Stepper Motor หยุด ทำงานหยุด สไลด์เข้า" THEN
       "Blackword SR(20)" := TRUE;   // SR flip-flop
   END_IF;
   IF "Output Step motor  Backword ทำงาน10" THEN "Blackword SR(20)" := FALSE; END_IF;
   #_w21 := "Blackword SR(20)";
   "Expected"(Expected1 := "Expected/Value_All".Expected_261,
              Expected2 := "Expected/Value_All".Expected_262,
              Expected3 := "Expected/Value_All".Expected_263,
              Expected4 := "Expected/Value_All".Expected_264,
              Expected5 := "Expected/Value_All".Expected_265,
              Expected6 := "Expected/Value_All".Expected_266,
              Expected7 := "Expected/Value_All".Expected_267,
              Expected8 := "Expected/Value_All".Expected_268,
              Expected9 := "Expected/Value_All".Expected_269,
              Expected10 := "Expected/Value_All".Expected_270,
              Expected11 := "Expected/Value_All".Expected_271,
              Expected12 := "Expected/Value_All".Expected_272,
              Expected13 := "Expected/Value_All".Expected_273,
              Expected14 := "Expected/Value_All".Expected_274,
              Expected15 := "Expected/Value_All".Expected_275,
              Expected16 := "Expected/Value_All".Expected_276,
              Expected17 := "Expected/Value_All".Expected_277,
              Expected18 := "Expected/Value_All".Expected_278,
              Expected19 := "Expected/Value_All".Expected_279,
              Expected20 := "Expected/Value_All".Expected_280,
              Expected21 := "Expected/Value_All".Expected_281,
              Expected22 := "Expected/Value_All".Expected_282,
              Expected23 := "Expected/Value_All".Expected_283,
              Expected24 := "Expected/Value_All".Expected_284,
              Expected25 := "Expected/Value_All".Expected_285,
              Expected26 := "Expected/Value_All".Expected_286,
              On_Motor => "Output Step Motor Blackword  No.11",
              ENO => #_w20);
   IF #_w20 AND "Output Step Motor Blackword  No.11" THEN
       "Blackword SR(21)" := TRUE;   // SR flip-flop
   END_IF;
   IF "Output Step motor  Backword ทำงาน11" THEN "Blackword SR(21)" := FALSE; END_IF;
   "IEC_Counter_0_DB_14".CTU(CU := "Blackword SR(21)" AND "Stepper Motor ทำงาน สไลด์เข้า",
                           R := "Output Step motor  Backword ทำงาน11",
                           PV := 2);
   IF "IEC_Counter_0_DB_14".Q AND "Stepper Motor หยุด ทำงานหยุด สไลด์เข้า" THEN
       "Blackword SR(22)" := TRUE;   // SR flip-flop
   END_IF;
   IF "Output Step motor  Backword ทำงาน11" THEN "Blackword SR(22)" := FALSE; END_IF;
   #_w23 := "Blackword SR(22)";
   "Expected"(Expected1 := "Expected/Value_All".Expected_287,
              Expected2 := "Expected/Value_All".Expected_288,
              Expected3 := "Expected/Value_All".Expected_289,
              Expected4 := "Expected/Value_All".Expected_290,
              Expected5 := "Expected/Value_All".Expected_291,
              Expected6 := "Expected/Value_All".Expected_292,
              Expected7 := "Expected/Value_All".Expected_293,
              Expected8 := "Expected/Value_All".Expected_294,
              Expected9 := "Expected/Value_All".Expected_295,
              Expected10 := "Expected/Value_All".Expected_296,
              Expected11 := "Expected/Value_All".Expected_297,
              Expected12 := "Expected/Value_All".Expected_298,
              Expected13 := "Expected/Value_All".Expected_299,
              Expected14 := "Expected/Value_All".Expected_300,
              Expected15 := "Expected/Value_All".Expected_301,
              Expected16 := "Expected/Value_All".Expected_302,
              Expected17 := "Expected/Value_All".Expected_303,
              Expected18 := "Expected/Value_All".Expected_304,
              Expected19 := "Expected/Value_All".Expected_305,
              Expected20 := "Expected/Value_All".Expected_306,
              Expected21 := "Expected/Value_All".Expected_307,
              Expected22 := "Expected/Value_All".Expected_308,
              Expected23 := "Expected/Value_All".Expected_309,
              Expected24 := "Expected/Value_All".Expected_310,
              Expected25 := "Expected/Value_All".Expected_311,
              Expected26 := "Expected/Value_All".Expected_312,
              On_Motor => "Output Step Motor Blackword  No.12",
              ENO => #_w22);
   IF #_w22 AND "Output Step Motor Blackword  No.12" THEN
       "Blackword SR(23)" := TRUE;   // SR flip-flop
   END_IF;
   IF "Output Step motor  Backword ทำงาน12" THEN "Blackword SR(23)" := FALSE; END_IF;
   "IEC_Counter_0_DB_15".CTU(CU := "Blackword SR(23)" AND "Stepper Motor ทำงาน สไลด์เข้า",
                           R := "Output Step motor  Backword ทำงาน12",
                           PV := 2);
   IF "IEC_Counter_0_DB_15".Q AND "Stepper Motor หยุด ทำงานหยุด สไลด์เข้า" THEN
       "Blackword SR(24)" := TRUE;   // SR flip-flop
   END_IF;
   IF "Output Step motor  Backword ทำงาน12" THEN "Blackword SR(24)" := FALSE; END_IF;
   #_w25 := "Blackword SR(24)";
   "Expected"(Expected1 := "Expected/Value_All".Expected_313,
              Expected2 := "Expected/Value_All".Expected_314,
              Expected3 := "Expected/Value_All".Expected_315,
              Expected4 := "Expected/Value_All".Expected_316,
              Expected5 := "Expected/Value_All".Expected_317,
              Expected6 := "Expected/Value_All".Expected_318,
              Expected7 := "Expected/Value_All".Expected_319,
              Expected8 := "Expected/Value_All".Expected_320,
              Expected9 := "Expected/Value_All".Expected_321,
              Expected10 := "Expected/Value_All".Expected_322,
              Expected11 := "Expected/Value_All".Expected_323,
              Expected12 := "Expected/Value_All".Expected_324,
              Expected13 := "Expected/Value_All".Expected_325,
              Expected14 := "Expected/Value_All".Expected_326,
              Expected15 := "Expected/Value_All".Expected_327,
              Expected16 := "Expected/Value_All".Expected_328,
              Expected17 := "Expected/Value_All".Expected_329,
              Expected18 := "Expected/Value_All".Expected_330,
              Expected19 := "Expected/Value_All".Expected_331,
              Expected20 := "Expected/Value_All".Expected_332,
              Expected21 := "Expected/Value_All".Expected_333,
              Expected22 := "Expected/Value_All".Expected_334,
              Expected23 := "Expected/Value_All".Expected_335,
              Expected24 := "Expected/Value_All".Expected_336,
              Expected25 := "Expected/Value_All".Expected_337,
              Expected26 := "Expected/Value_All".Expected_338,
              On_Motor => "Output Step Motor Blackword  No.13",
              ENO => #_w24);
   IF #_w24 AND "Output Step Motor Blackword  No.13" THEN
       "Blackword SR(25)" := TRUE;   // SR flip-flop
   END_IF;
   IF "Output Step motor  Backword ทำงาน13" THEN "Blackword SR(25)" := FALSE; END_IF;
   "IEC_Counter_0_DB_16".CTU(CU := "Blackword SR(25)" AND "Stepper Motor ทำงาน สไลด์เข้า",
                           R := "Output Step motor  Backword ทำงาน13",
                           PV := 2);
   IF "IEC_Counter_0_DB_16".Q AND "Stepper Motor หยุด ทำงานหยุด สไลด์เข้า" THEN
       "Blackword SR(26)" := TRUE;   // SR flip-flop
   END_IF;
   IF "Output Step motor  Backword ทำงาน13" THEN "Blackword SR(26)" := FALSE; END_IF;
   #_w27 := "Blackword SR(26)";
   "Expected"(Expected1 := "Expected/Value_All".Expected_339,
              Expected2 := "Expected/Value_All".Expected_340,
              Expected3 := "Expected/Value_All".Expected_341,
              Expected4 := "Expected/Value_All".Expected_342,
              Expected5 := "Expected/Value_All".Expected_343,
              Expected6 := "Expected/Value_All".Expected_344,
              Expected7 := "Expected/Value_All".Expected_345,
              Expected8 := "Expected/Value_All".Expected_346,
              Expected9 := "Expected/Value_All".Expected_347,
              Expected10 := "Expected/Value_All".Expected_348,
              Expected11 := "Expected/Value_All".Expected_349,
              Expected12 := "Expected/Value_All".Expected_350,
              Expected13 := "Expected/Value_All".Expected_351,
              Expected14 := "Expected/Value_All".Expected_352,
              Expected15 := "Expected/Value_All".Expected_353,
              Expected16 := "Expected/Value_All".Expected_354,
              Expected17 := "Expected/Value_All".Expected_355,
              Expected18 := "Expected/Value_All".Expected_356,
              Expected19 := "Expected/Value_All".Expected_357,
              Expected20 := "Expected/Value_All".Expected_358,
              Expected21 := "Expected/Value_All".Expected_359,
              Expected22 := "Expected/Value_All".Expected_360,
              Expected23 := "Expected/Value_All".Expected_361,
              Expected24 := "Expected/Value_All".Expected_362,
              Expected25 := "Expected/Value_All".Expected_363,
              Expected26 := "Expected/Value_All".Expected_364,
              On_Motor => "Output Step Motor Blackword  No.14",
              ENO => #_w26);
   IF #_w26 AND "Output Step Motor Blackword  No.14" THEN
       "Blackword SR(27)" := TRUE;   // SR flip-flop
   END_IF;
   IF "Output Step motor  Backword ทำงาน14" THEN "Blackword SR(27)" := FALSE; END_IF;
   "IEC_Counter_0_DB_17".CTU(CU := "Blackword SR(27)" AND "Stepper Motor ทำงาน สไลด์เข้า",
                           R := "Output Step motor  Backword ทำงาน14",
                           PV := 2);
   IF "IEC_Counter_0_DB_17".Q AND "Stepper Motor หยุด ทำงานหยุด สไลด์เข้า" THEN
       "Blackword SR(28)" := TRUE;   // SR flip-flop
   END_IF;
   IF "Output Step motor  Backword ทำงาน14" THEN "Blackword SR(28)" := FALSE; END_IF;
   #_w29 := "Blackword SR(28)";
   "Expected"(Expected1 := "Expected/Value_All".Expected_365,
              Expected2 := "Expected/Value_All".Expected_366,
              Expected3 := "Expected/Value_All".Expected_367,
              Expected4 := "Expected/Value_All".Expected_368,
              Expected5 := "Expected/Value_All".Expected_369,
              Expected6 := "Expected/Value_All".Expected_370,
              Expected7 := "Expected/Value_All".Expected_371,
              Expected8 := "Expected/Value_All".Expected_372,
              Expected9 := "Expected/Value_All".Expected_373,
              Expected10 := "Expected/Value_All".Expected_374,
              Expected11 := "Expected/Value_All".Expected_375,
              Expected12 := "Expected/Value_All".Expected_376,
              Expected13 := "Expected/Value_All".Expected_377,
              Expected14 := "Expected/Value_All".Expected_378,
              Expected15 := "Expected/Value_All".Expected_379,
              Expected16 := "Expected/Value_All".Expected_380,
              Expected17 := "Expected/Value_All".Expected_381,
              Expected18 := "Expected/Value_All".Expected_382,
              Expected19 := "Expected/Value_All".Expected_383,
              Expected20 := "Expected/Value_All".Expected_384,
              Expected21 := "Expected/Value_All".Expected_385,
              Expected22 := "Expected/Value_All".Expected_386,
              Expected23 := "Expected/Value_All".Expected_387,
              Expected24 := "Expected/Value_All".Expected_388,
              Expected25 := "Expected/Value_All".Expected_389,
              Expected26 := "Expected/Value_All".Expected_390,
              On_Motor => "Output Step Motor Blackword  No.15",
              ENO => #_w28);
   IF #_w28 AND "Output Step Motor Blackword  No.15" THEN
       "Blackword SR(29)" := TRUE;   // SR flip-flop
   END_IF;
   IF "Output Step motor  Backword ทำงาน15" THEN "Blackword SR(29)" := FALSE; END_IF;
   "IEC_Counter_0_DB_18".CTU(CU := "Blackword SR(29)" AND "Stepper Motor ทำงาน สไลด์เข้า",
                           R := "Output Step motor  Backword ทำงาน15",
                           PV := 2);
   IF "IEC_Counter_0_DB_18".Q AND "Stepper Motor หยุด ทำงานหยุด สไลด์เข้า" THEN
       "Blackword SR(30)" := TRUE;   // SR flip-flop
   END_IF;
   IF "Output Step motor  Backword ทำงาน15" THEN "Blackword SR(30)" := FALSE; END_IF;
   #_w31 := "Blackword SR(30)";
   "Expected"(Expected1 := "Expected/Value_All".Expected_391,
              Expected2 := "Expected/Value_All".Expected_392,
              Expected3 := "Expected/Value_All".Expected_393,
              Expected4 := "Expected/Value_All".Expected_394,
              Expected5 := "Expected/Value_All".Expected_395,
              Expected6 := "Expected/Value_All".Expected_396,
              Expected7 := "Expected/Value_All".Expected_397,
              Expected8 := "Expected/Value_All".Expected_398,
              Expected9 := "Expected/Value_All".Expected_399,
              Expected10 := "Expected/Value_All".Expected_400,
              Expected11 := "Expected/Value_All".Expected_401,
              Expected12 := "Expected/Value_All".Expected_402,
              Expected13 := "Expected/Value_All".Expected_403,
              Expected14 := "Expected/Value_All".Expected_404,
              Expected15 := "Expected/Value_All".Expected_405,
              Expected16 := "Expected/Value_All".Expected_406,
              Expected17 := "Expected/Value_All".Expected_407,
              Expected18 := "Expected/Value_All".Expected_408,
              Expected19 := "Expected/Value_All".Expected_409,
              Expected20 := "Expected/Value_All".Expected_410,
              Expected21 := "Expected/Value_All".Expected_411,
              Expected22 := "Expected/Value_All".Expected_412,
              Expected23 := "Expected/Value_All".Expected_413,
              Expected24 := "Expected/Value_All".Expected_414,
              Expected25 := "Expected/Value_All".Expected_415,
              Expected26 := "Expected/Value_All".Expected_416,
              On_Motor => "Output Step Motor Blackword  No.16",
              ENO => #_w30);
   IF #_w30 AND "Output Step Motor Blackword  No.16" THEN
       "Blackword SR(31)" := TRUE;   // SR flip-flop
   END_IF;
   IF "Output Step motor  Backword ทำงาน16" THEN "Blackword SR(31)" := FALSE; END_IF;
   "IEC_Counter_0_DB_19".CTU(CU := "Blackword SR(31)" AND "Stepper Motor ทำงาน สไลด์เข้า",
                           R := "Output Step motor  Backword ทำงาน16",
                           PV := 2);
   IF "IEC_Counter_0_DB_19".Q AND "Stepper Motor หยุด ทำงานหยุด สไลด์เข้า" THEN
       "Blackword SR(32)" := TRUE;   // SR flip-flop
   END_IF;
   IF "Output Step motor  Backword ทำงาน16" THEN "Blackword SR(32)" := FALSE; END_IF;
   #_w33 := "Blackword SR(32)";
   "Expected"(Expected1 := "Expected/Value_All".Expected_417,
              Expected2 := "Expected/Value_All".Expected_418,
              Expected3 := "Expected/Value_All".Expected_419,
              Expected4 := "Expected/Value_All".Expected_420,
              Expected5 := "Expected/Value_All".Expected_421,
              Expected6 := "Expected/Value_All".Expected_422,
              Expected7 := "Expected/Value_All".Expected_423,
              Expected8 := "Expected/Value_All".Expected_424,
              Expected9 := "Expected/Value_All".Expected_425,
              Expected10 := "Expected/Value_All".Expected_426,
              Expected11 := "Expected/Value_All".Expected_427,
              Expected12 := "Expected/Value_All".Expected_428,
              Expected13 := "Expected/Value_All".Expected_429,
              Expected14 := "Expected/Value_All".Expected_430,
              Expected15 := "Expected/Value_All".Expected_431,
              Expected16 := "Expected/Value_All".Expected_432,
              Expected17 := "Expected/Value_All".Expected_433,
              Expected18 := "Expected/Value_All".Expected_434,
              Expected19 := "Expected/Value_All".Expected_435,
              Expected20 := "Expected/Value_All".Expected_436,
              Expected21 := "Expected/Value_All".Expected_437,
              Expected22 := "Expected/Value_All".Expected_438,
              Expected23 := "Expected/Value_All".Expected_439,
              Expected24 := "Expected/Value_All".Expected_440,
              Expected25 := "Expected/Value_All".Expected_441,
              Expected26 := "Expected/Value_All".Expected_442,
              On_Motor => "Output Step Motor Blackword  No.17",
              ENO => #_w32);
   IF #_w32 AND "Output Step Motor Blackword  No.17" THEN
       "Blackword SR(33)" := TRUE;   // SR flip-flop
   END_IF;
   IF "Output Step motor  Backword ทำงาน17" THEN "Blackword SR(33)" := FALSE; END_IF;
   "IEC_Counter_0_DB_20".CTU(CU := "Blackword SR(33)" AND "Stepper Motor ทำงาน สไลด์เข้า",
                           R := "Output Step motor  Backword ทำงาน17",
                           PV := 2);
   IF "IEC_Counter_0_DB_20".Q AND "Stepper Motor หยุด ทำงานหยุด สไลด์เข้า" THEN
       "Blackword SR(34)" := TRUE;   // SR flip-flop
   END_IF;
   IF "Output Step motor  Backword ทำงาน17" THEN "Blackword SR(34)" := FALSE; END_IF;
   #_w35 := "Blackword SR(34)";
   "Expected"(Expected1 := "Expected/Value_All".Expected_443,
              Expected2 := "Expected/Value_All".Expected_444,
              Expected3 := "Expected/Value_All".Expected_445,
              Expected4 := "Expected/Value_All".Expected_446,
              Expected5 := "Expected/Value_All".Expected_447,
              Expected6 := "Expected/Value_All".Expected_448,
              Expected7 := "Expected/Value_All".Expected_449,
              Expected8 := "Expected/Value_All".Expected_450,
              Expected9 := "Expected/Value_All".Expected_451,
              Expected10 := "Expected/Value_All".Expected_452,
              Expected11 := "Expected/Value_All".Expected_453,
              Expected12 := "Expected/Value_All".Expected_454,
              Expected13 := "Expected/Value_All".Expected_455,
              Expected14 := "Expected/Value_All".Expected_456,
              Expected15 := "Expected/Value_All".Expected_457,
              Expected16 := "Expected/Value_All".Expected_458,
              Expected17 := "Expected/Value_All".Expected_459,
              Expected18 := "Expected/Value_All".Expected_460,
              Expected19 := "Expected/Value_All".Expected_461,
              Expected20 := "Expected/Value_All".Expected_462,
              Expected21 := "Expected/Value_All".Expected_463,
              Expected22 := "Expected/Value_All".Expected_464,
              Expected23 := "Expected/Value_All".Expected_465,
              Expected24 := "Expected/Value_All".Expected_466,
              Expected25 := "Expected/Value_All".Expected_467,
              Expected26 := "Expected/Value_All".Expected_468,
              On_Motor => "Output Step Motor Blackword  No.18",
              ENO => #_w34);
   IF #_w34 AND "Output Step Motor Blackword  No.18" THEN
       "Blackword SR(35)" := TRUE;   // SR flip-flop
   END_IF;
   IF "Output Step motor  Backword ทำงาน18" THEN "Blackword SR(35)" := FALSE; END_IF;
   "IEC_Counter_0_DB_21".CTU(CU := "Blackword SR(35)" AND "Stepper Motor ทำงาน สไลด์เข้า",
                           R := "Output Step motor  Backword ทำงาน18",
                           PV := 2);
   IF "IEC_Counter_0_DB_21".Q AND "Stepper Motor หยุด ทำงานหยุด สไลด์เข้า" THEN
       "Blackword SR(36)" := TRUE;   // SR flip-flop
   END_IF;
   IF "Output Step motor  Backword ทำงาน18" THEN "Blackword SR(36)" := FALSE; END_IF;
   #_w37 := "Blackword SR(36)";
   "Expected"(Expected1 := "Expected/Value_All".Expected_469,
              Expected2 := "Expected/Value_All".Expected_470,
              Expected3 := "Expected/Value_All".Expected_471,
              Expected4 := "Expected/Value_All".Expected_472,
              Expected5 := "Expected/Value_All".Expected_473,
              Expected6 := "Expected/Value_All".Expected_474,
              Expected7 := "Expected/Value_All".Expected_475,
              Expected8 := "Expected/Value_All".Expected_476,
              Expected9 := "Expected/Value_All".Expected_477,
              Expected10 := "Expected/Value_All".Expected_478,
              Expected11 := "Expected/Value_All".Expected_479,
              Expected12 := "Expected/Value_All".Expected_480,
              Expected13 := "Expected/Value_All".Expected_481,
              Expected14 := "Expected/Value_All".Expected_482,
              Expected15 := "Expected/Value_All".Expected_483,
              Expected16 := "Expected/Value_All".Expected_484,
              Expected17 := "Expected/Value_All".Expected_485,
              Expected18 := "Expected/Value_All".Expected_486,
              Expected19 := "Expected/Value_All".Expected_487,
              Expected20 := "Expected/Value_All".Expected_488,
              Expected21 := "Expected/Value_All".Expected_489,
              Expected22 := "Expected/Value_All".Expected_490,
              Expected23 := "Expected/Value_All".Expected_491,
              Expected24 := "Expected/Value_All".Expected_492,
              Expected25 := "Expected/Value_All".Expected_493,
              Expected26 := "Expected/Value_All".Expected_494,
              On_Motor => "Output Step Motor Blackword  No.19",
              ENO => #_w36);
   IF #_w36 AND "Output Step Motor Blackword  No.19" THEN
       "Blackword SR(37)" := TRUE;   // SR flip-flop
   END_IF;
   IF "Output Step motor  Backword ทำงาน19" THEN "Blackword SR(37)" := FALSE; END_IF;
   "IEC_Counter_0_DB_22".CTU(CU := "Blackword SR(37)" AND "Stepper Motor ทำงาน สไลด์เข้า",
                           R := "Output Step motor  Backword ทำงาน19",
                           PV := 2);
   IF "IEC_Counter_0_DB_22".Q AND "Stepper Motor หยุด ทำงานหยุด สไลด์เข้า" THEN
       "Blackword SR(38)" := TRUE;   // SR flip-flop
   END_IF;
   IF "Output Step motor  Backword ทำงาน19" THEN "Blackword SR(38)" := FALSE; END_IF;
   #_w39 := "Blackword SR(38)";
   "Expected"(Expected1 := "Expected/Value_All".Expected_495,
              Expected2 := "Expected/Value_All".Expected_496,
              Expected3 := "Expected/Value_All".Expected_497,
              Expected4 := "Expected/Value_All".Expected_498,
              Expected5 := "Expected/Value_All".Expected_499,
              Expected6 := "Expected/Value_All".Expected_500,
              Expected7 := "Expected/Value_All".Expected_501,
              Expected8 := "Expected/Value_All".Expected_502,
              Expected9 := "Expected/Value_All".Expected_503,
              Expected10 := "Expected/Value_All".Expected_504,
              Expected11 := "Expected/Value_All".Expected_505,
              Expected12 := "Expected/Value_All".Expected_506,
              Expected13 := "Expected/Value_All".Expected_507,
              Expected14 := "Expected/Value_All".Expected_508,
              Expected15 := "Expected/Value_All".Expected_509,
              Expected16 := "Expected/Value_All".Expected_510,
              Expected17 := "Expected/Value_All".Expected_511,
              Expected18 := "Expected/Value_All".Expected_512,
              Expected19 := "Expected/Value_All".Expected_513,
              Expected20 := "Expected/Value_All".Expected_514,
              Expected21 := "Expected/Value_All".Expected_515,
              Expected22 := "Expected/Value_All".Expected_516,
              Expected23 := "Expected/Value_All".Expected_517,
              Expected24 := "Expected/Value_All".Expected_518,
              Expected25 := "Expected/Value_All".Expected_519,
              Expected26 := "Expected/Value_All".Expected_520,
              On_Motor => "Output Step Motor Blackword  No.20",
              ENO => #_w38);
   IF #_w38 AND "Output Step Motor Blackword  No.20" THEN
       "Blackword SR(39)" := TRUE;   // SR flip-flop
   END_IF;
   IF "Output Step motor  Backword ทำงาน20" THEN "Blackword SR(39)" := FALSE; END_IF;
   "IEC_Counter_0_DB_23".CTU(CU := "Blackword SR(39)" AND "Stepper Motor ทำงาน สไลด์เข้า",
                           R := "Output Step motor  Backword ทำงาน20",
                           PV := 2);
   IF "IEC_Counter_0_DB_23".Q AND "Stepper Motor หยุด ทำงานหยุด สไลด์เข้า" THEN
       "Blackword SR(40)" := TRUE;   // SR flip-flop
   END_IF;
   IF "Output Step motor  Backword ทำงาน20" THEN "Blackword SR(40)" := FALSE; END_IF;
   #"Step motor  Backword ทำงาน" := #_w3 OR #_w5 OR #_w7 OR #_w9 OR #_w11 OR #_w13 OR #_w15 OR #_w17 OR #_w19 OR #_w21 OR #_w23 OR #_w25 OR #_w27 OR #_w29 OR #_w31 OR #_w33 OR #_w35 OR #_w37 OR #_w39 OR "Blackword SR(40)";
   "IEC_Timer_0_DB_2".TONR(IN := #"Step motor  Backword ทำงาน",
                           R := NOT #"Step motor  Backword ทำงาน",
                           PT := #"เวลาเคลื่อนที่ของ Stepper Motor1จาก Box1_Backword");
   "Output Step motor  Backword ทำงาน1" := "IEC_Timer_0_DB_2".Q OR "มีการปุ่มกดยืนยัน";
   "IEC_Timer_0_DB_3".TONR(IN := #"Step motor  Backword ทำงาน",
                           R := NOT #"Step motor  Backword ทำงาน",
                           PT := #"เวลาเคลื่อนที่ของ Stepper Motor1จาก Box2_Backword");
   "Output Step motor  Backword ทำงาน2" := "IEC_Timer_0_DB_3".Q OR "มีการปุ่มกดยืนยัน";
   "IEC_Timer_0_DB_35".TONR(IN := #"Step motor  Backword ทำงาน",
                           R := NOT #"Step motor  Backword ทำงาน",
                           PT := #"เวลาเคลื่อนที่ของ Stepper Motor1จาก Box2_Backword");
   "Output Step motor  Backword ทำงาน3" := "IEC_Timer_0_DB_35".Q OR "มีการปุ่มกดยืนยัน";
   "IEC_Timer_0_DB_37".TONR(IN := #"Step motor  Backword ทำงาน",
                           R := NOT #"Step motor  Backword ทำงาน",
                           PT := #"เวลาเคลื่อนที่ของ Stepper Motor1จาก Box2_Backword");
   "Output Step motor  Backword ทำงาน4" := "IEC_Timer_0_DB_37".Q OR "มีการปุ่มกดยืนยัน";
   "IEC_Timer_0_DB_38".TONR(IN := #"Step motor  Backword ทำงาน",
                           R := NOT #"Step motor  Backword ทำงาน",
                           PT := #"เวลาเคลื่อนที่ของ Stepper Motor1จาก Box2_Backword");
   "Output Step motor  Backword ทำงาน5" := "IEC_Timer_0_DB_38".Q OR "มีการปุ่มกดยืนยัน";
   "IEC_Timer_0_DB_39".TONR(IN := #"Step motor  Backword ทำงาน",
                           R := NOT #"Step motor  Backword ทำงาน",
                           PT := #"เวลาเคลื่อนที่ของ Stepper Motor1จาก Box2_Backword");
   "Output Step motor  Backword ทำงาน6" := "IEC_Timer_0_DB_39".Q OR "มีการปุ่มกดยืนยัน";
   "IEC_Timer_0_DB_40".TONR(IN := #"Step motor  Backword ทำงาน",
                           R := NOT #"Step motor  Backword ทำงาน",
                           PT := #"เวลาเคลื่อนที่ของ Stepper Motor1จาก Box2_Backword");
   "Output Step motor  Backword ทำงาน7" := "IEC_Timer_0_DB_40".Q OR "มีการปุ่มกดยืนยัน";
   "IEC_Timer_0_DB_41".TONR(IN := #"Step motor  Backword ทำงาน",
                           R := NOT #"Step motor  Backword ทำงาน",
                           PT := #"เวลาเคลื่อนที่ของ Stepper Motor1จาก Box2_Backword");
   "Output Step motor  Backword ทำงาน8" := "IEC_Timer_0_DB_41".Q OR "มีการปุ่มกดยืนยัน";
   "IEC_Timer_0_DB_42".TONR(IN := #"Step motor  Backword ทำงาน",
                           R := NOT #"Step motor  Backword ทำงาน",
                           PT := #"เวลาเคลื่อนที่ของ Stepper Motor1จาก Box2_Backword");
   "Output Step motor  Backword ทำงาน9" := "IEC_Timer_0_DB_42".Q OR "มีการปุ่มกดยืนยัน";
   "IEC_Timer_0_DB_43".TONR(IN := #"Step motor  Backword ทำงาน",
                           R := NOT #"Step motor  Backword ทำงาน",
                           PT := #"เวลาเคลื่อนที่ของ Stepper Motor1จาก Box2_Backword");
   "Output Step motor  Backword ทำงาน10" := "IEC_Timer_0_DB_43".Q OR "มีการปุ่มกดยืนยัน";
   "IEC_Timer_0_DB_44".TONR(IN := #"Step motor  Backword ทำงาน",
                           R := NOT #"Step motor  Backword ทำงาน",
                           PT := #"เวลาเคลื่อนที่ของ Stepper Motor1จาก Box2_Backword");
   "Output Step motor  Backword ทำงาน11" := "IEC_Timer_0_DB_44".Q OR "มีการปุ่มกดยืนยัน";
   "IEC_Timer_0_DB_45".TONR(IN := #"Step motor  Backword ทำงาน",
                           R := NOT #"Step motor  Backword ทำงาน",
                           PT := #"เวลาเคลื่อนที่ของ Stepper Motor1จาก Box2_Backword");
   "Output Step motor  Backword ทำงาน12" := "IEC_Timer_0_DB_45".Q OR "มีการปุ่มกดยืนยัน";
   "IEC_Timer_0_DB_46".TONR(IN := #"Step motor  Backword ทำงาน",
                           R := NOT #"Step motor  Backword ทำงาน",
                           PT := #"เวลาเคลื่อนที่ของ Stepper Motor1จาก Box2_Backword");
   "Output Step motor  Backword ทำงาน13" := "IEC_Timer_0_DB_46".Q OR "มีการปุ่มกดยืนยัน";
   "IEC_Timer_0_DB_47".TONR(IN := #"Step motor  Backword ทำงาน",
                           R := NOT #"Step motor  Backword ทำงาน",
                           PT := #"เวลาเคลื่อนที่ของ Stepper Motor1จาก Box2_Backword");
   "Output Step motor  Backword ทำงาน14" := "IEC_Timer_0_DB_47".Q OR "มีการปุ่มกดยืนยัน";
   "IEC_Timer_0_DB_48".TONR(IN := #"Step motor  Backword ทำงาน",
                           R := NOT #"Step motor  Backword ทำงาน",
                           PT := #"เวลาเคลื่อนที่ของ Stepper Motor1จาก Box2_Backword");
   "Output Step motor  Backword ทำงาน15" := "IEC_Timer_0_DB_48".Q OR "มีการปุ่มกดยืนยัน";
   "IEC_Timer_0_DB_49".TONR(IN := #"Step motor  Backword ทำงาน",
                           R := NOT #"Step motor  Backword ทำงาน",
                           PT := #"เวลาเคลื่อนที่ของ Stepper Motor1จาก Box2_Backword");
   "Output Step motor  Backword ทำงาน16" := "IEC_Timer_0_DB_49".Q OR "มีการปุ่มกดยืนยัน";
   "IEC_Timer_0_DB_50".TONR(IN := #"Step motor  Backword ทำงาน",
                           R := NOT #"Step motor  Backword ทำงาน",
                           PT := #"เวลาเคลื่อนที่ของ Stepper Motor1จาก Box2_Backword");
   "Output Step motor  Backword ทำงาน17" := "IEC_Timer_0_DB_50".Q OR "มีการปุ่มกดยืนยัน";
   "IEC_Timer_0_DB_51".TONR(IN := #"Step motor  Backword ทำงาน",
                           R := NOT #"Step motor  Backword ทำงาน",
                           PT := #"เวลาเคลื่อนที่ของ Stepper Motor1จาก Box2_Backword");
   "Output Step motor  Backword ทำงาน18" := "IEC_Timer_0_DB_51".Q OR "มีการปุ่มกดยืนยัน";
   "IEC_Timer_0_DB_52".TONR(IN := #"Step motor  Backword ทำงาน",
                           R := NOT #"Step motor  Backword ทำงาน",
                           PT := #"เวลาเคลื่อนที่ของ Stepper Motor1จาก Box2_Backword");
   "Output Step motor  Backword ทำงาน19" := "IEC_Timer_0_DB_52".Q OR "มีการปุ่มกดยืนยัน";
   "IEC_Timer_0_DB_53".TONR(IN := #"Step motor  Backword ทำงาน",
                           R := NOT #"Step motor  Backword ทำงาน",
                           PT := #"เวลาเคลื่อนที่ของ Stepper Motor1จาก Box2_Backword");
   "Output Step motor  Backword ทำงาน20" := "IEC_Timer_0_DB_53".Q OR "มีการปุ่มกดยืนยัน";
END_REGION
END_FUNCTION_BLOCK

// folder: System_In(จัดเก็บ)/Step motor No.3

FUNCTION_BLOCK "Step motor ซ้าน-ขวา ตามแกน X  No.1_Forword"   // FB3, LAD
{ S7_Optimized_Access := 'TRUE' }
VERSION : 0.1
   VAR_INPUT
      "TIME ที่ใช้ไป แกน X.1" : Time;
      "TIME ที่ใช้ไป แกน X.2" : Time;
      "TIME ที่ใช้ไป แกน X.3" : Time;
      "TIME ที่ใช้ไป แกน X.4" : Time;
      "TIME ที่ใช้ไป แกน X.5" : Time;
      "TIME ที่ใช้ไป แกน X.6" : Time;
      "TIME ที่ใช้ไป แกน X.7" : Time;
      "TIME ที่ใช้ไป แกน X.8" : Time;
      "TIME ที่ใช้ไป แกน X.9" : Time;
      "TIME ที่ใช้ไป แกน X.10" : Time;
      "TIME ที่ใช้ไป แกน X.11" : Time;
      "TIME ที่ใช้ไป แกน X.12" : Time;
      "TIME ที่ใช้ไป แกน X.13" : Time;
      "TIME ที่ใช้ไป แกน X.14" : Time;
      "TIME ที่ใช้ไป แกน X.15" : Time;
      "TIME ที่ใช้ไป แกน X.16" : Time;
      "TIME ที่ใช้ไป แกน X.17" : Time;
      "TIME ที่ใช้ไป แกน X.18" : Time;
      "TIME ที่ใช้ไป แกน X.19" : Time;
      "TIME ที่ใช้ไป แกน X.20" : Time;
      "TIME ที่ใช้ไป แกน X.21" : Time;
      "TIME ที่ใช้ไป แกน X.22" : Time;
      "TIME ที่ใช้ไป แกน X.23" : Time;
      "TIME ที่ใช้ไป แกน X.24" : Time;
      "TIME ที่ใช้ไป แกน X.25" : Time;
      "TIME ที่ใช้ไป แกน X.26" : Time;
   END_VAR
   VAR_IN_OUT
      "Stepper Motor  ทำงาน3" : Bool;
   END_VAR
   VAR_TEMP   // added for the SCL form of the ladder/FBD networks
      _w1 : Bool;
      _w2 : Bool;
      _w3 : Bool;
      _w4 : Bool;
      _w5 : Bool;
      _w6 : Bool;
      _w7 : Bool;
      _w8 : Bool;
      _w9 : Bool;
      _w10 : Bool;
      _w11 : Bool;
      _w12 : Bool;
      _w13 : Bool;
      _w14 : Bool;
      _w15 : Bool;
      _w16 : Bool;
      _w17 : Bool;
      _w18 : Bool;
      _w19 : Bool;
      _w20 : Bool;
      _w21 : Bool;
      _w22 : Bool;
      _w23 : Bool;
      _w24 : Bool;
      _w25 : Bool;
      _w26 : Bool;
      _w27 : Bool;
      _w28 : Bool;
      _w29 : Bool;
      _w30 : Bool;
      _w31 : Bool;
      _w32 : Bool;
      _w33 : Bool;
      _w34 : Bool;
      _w35 : Bool;
      _w36 : Bool;
      _w37 : Bool;
      _w38 : Bool;
      _w39 : Bool;
      _w40 : Bool;
      _w41 : Bool;
      _w42 : Bool;
      _w43 : Bool;
      _w44 : Bool;
      _w45 : Bool;
      _w46 : Bool;
      _w47 : Bool;
      _w48 : Bool;
      _w49 : Bool;
      _w50 : Bool;
      _w51 : Bool;
   END_VAR
BEGIN

REGION Network 1
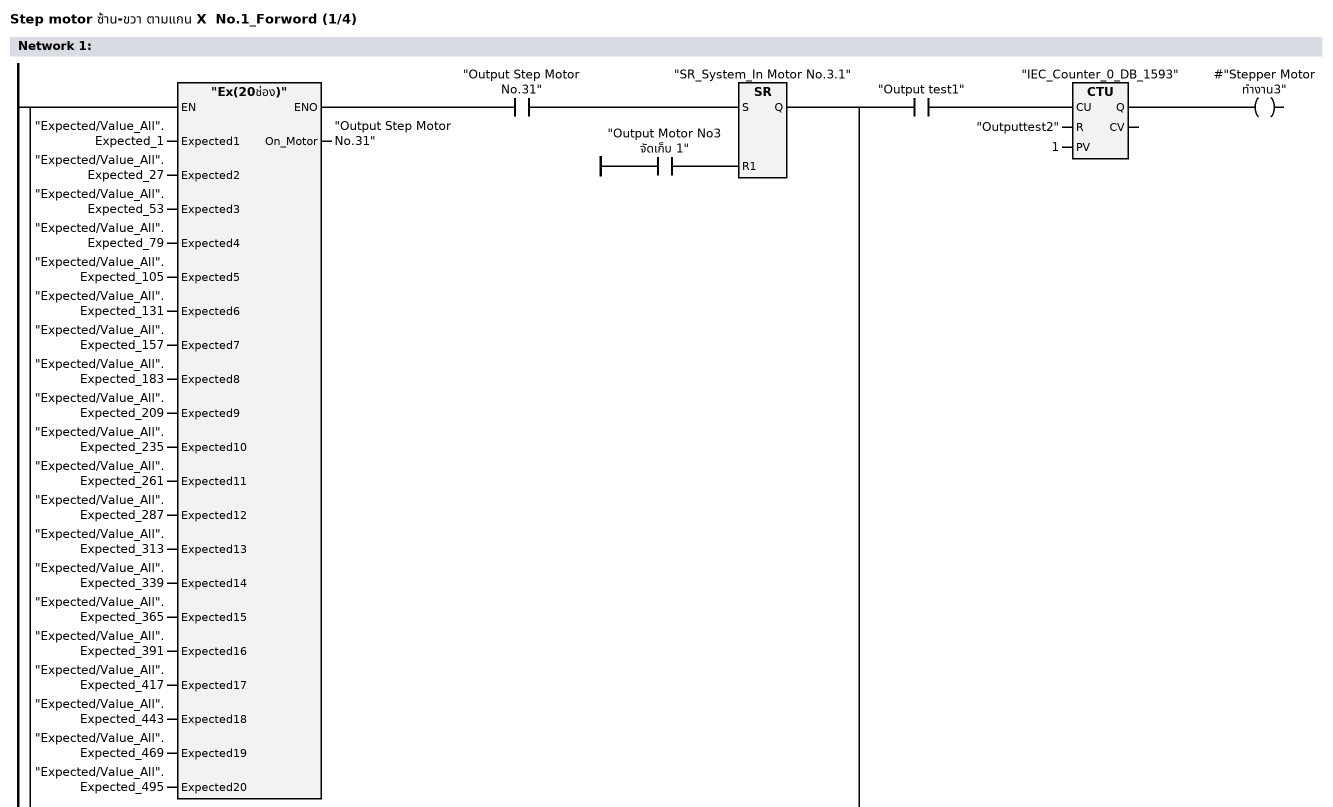
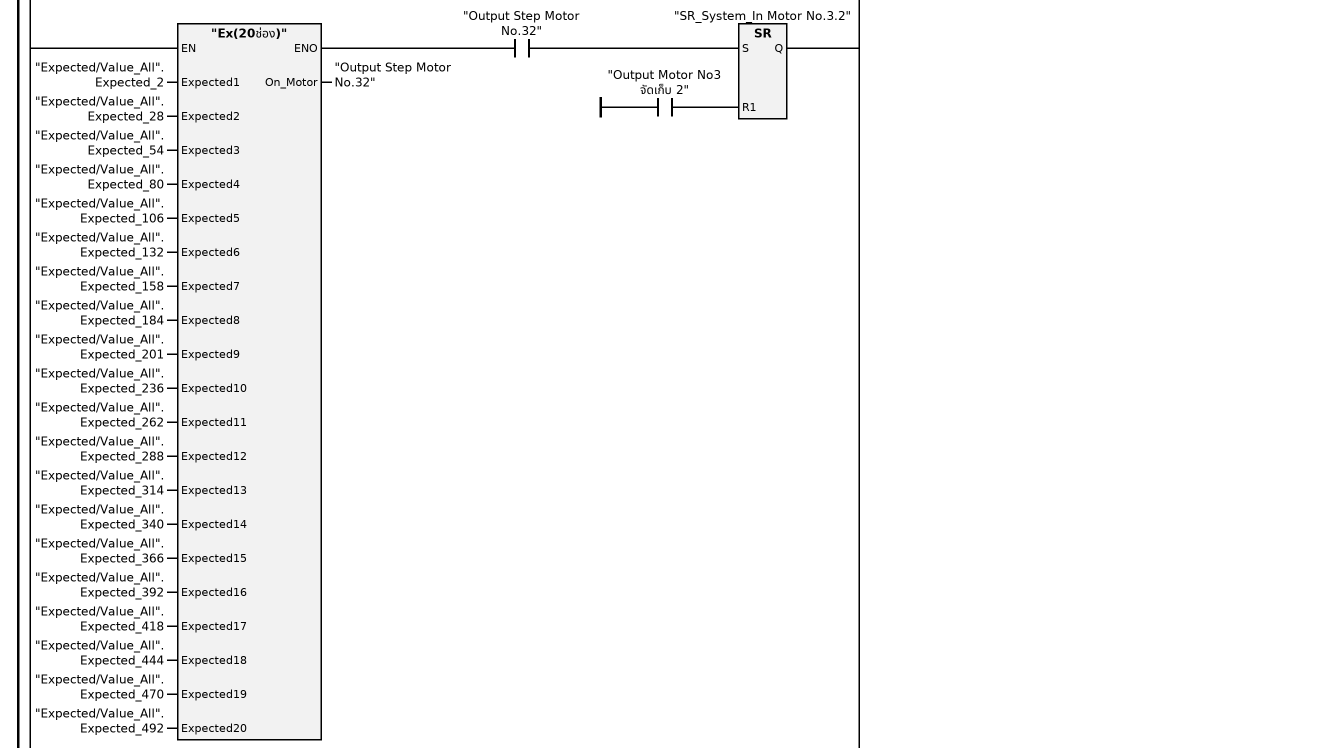
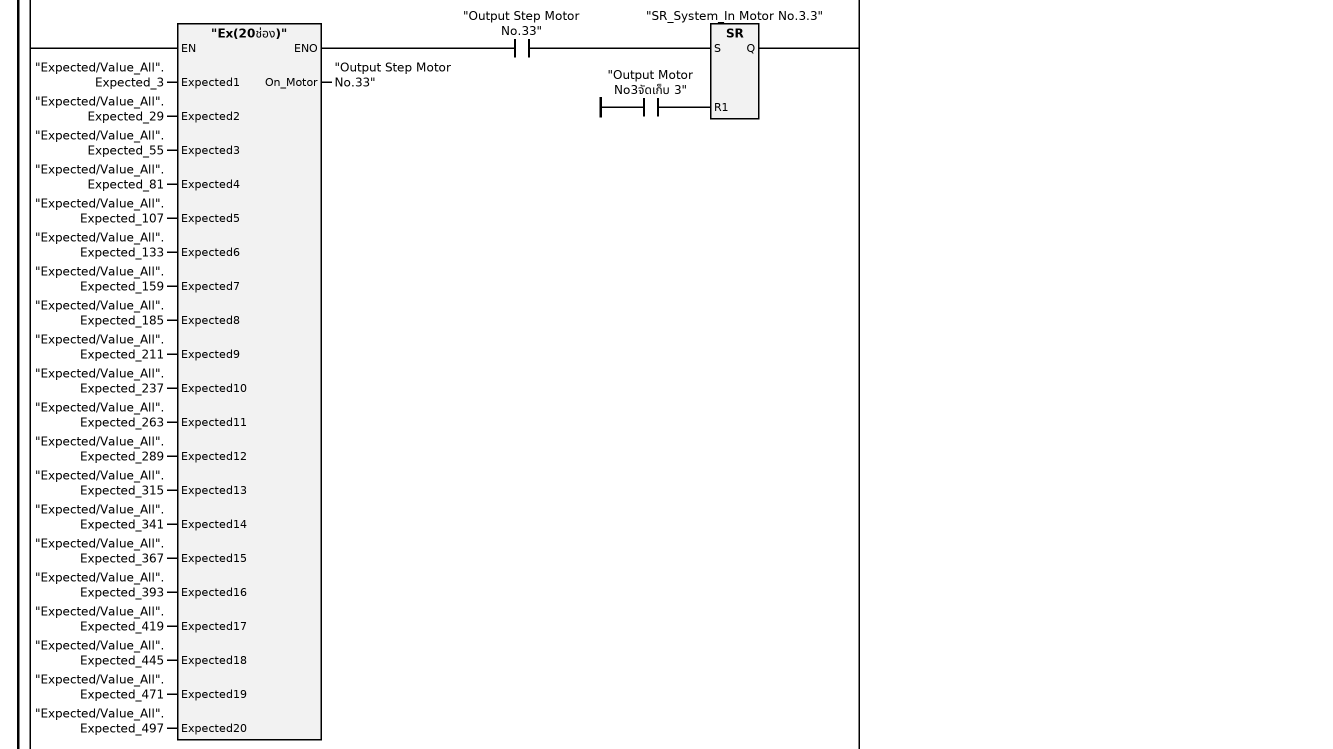
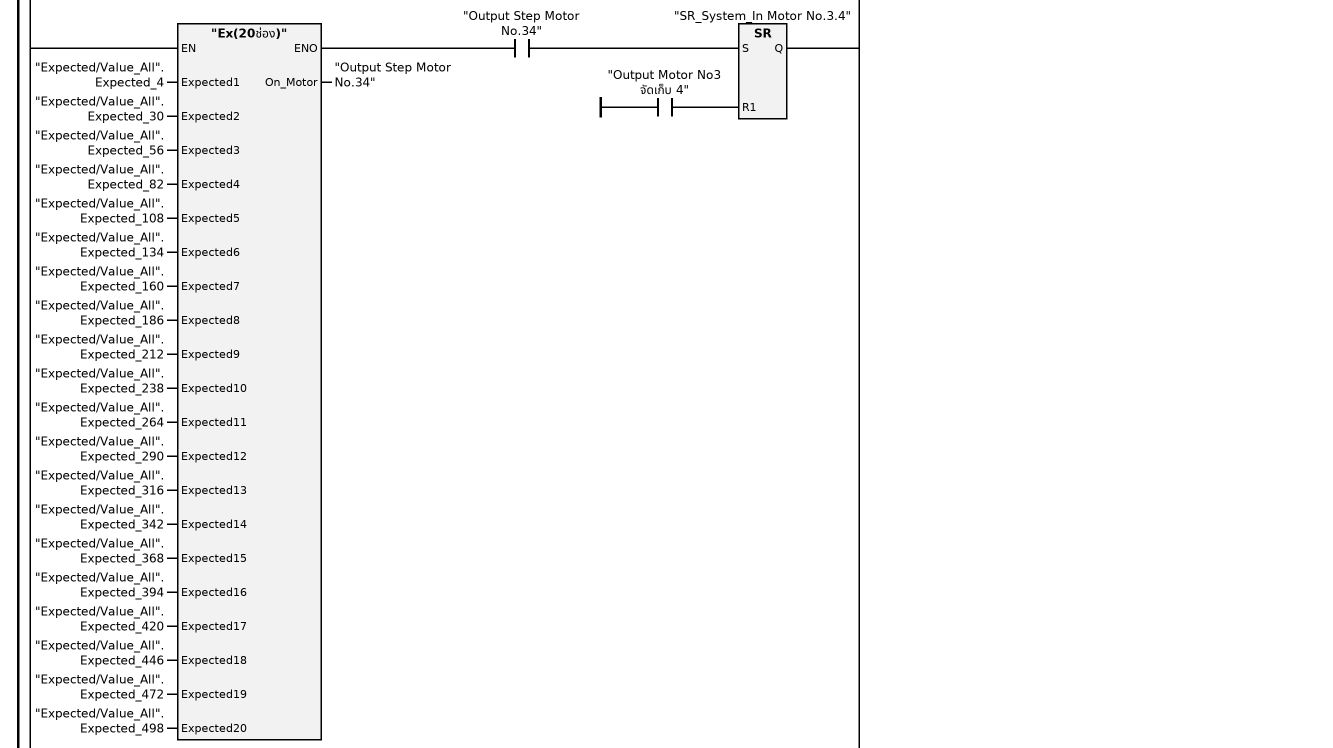
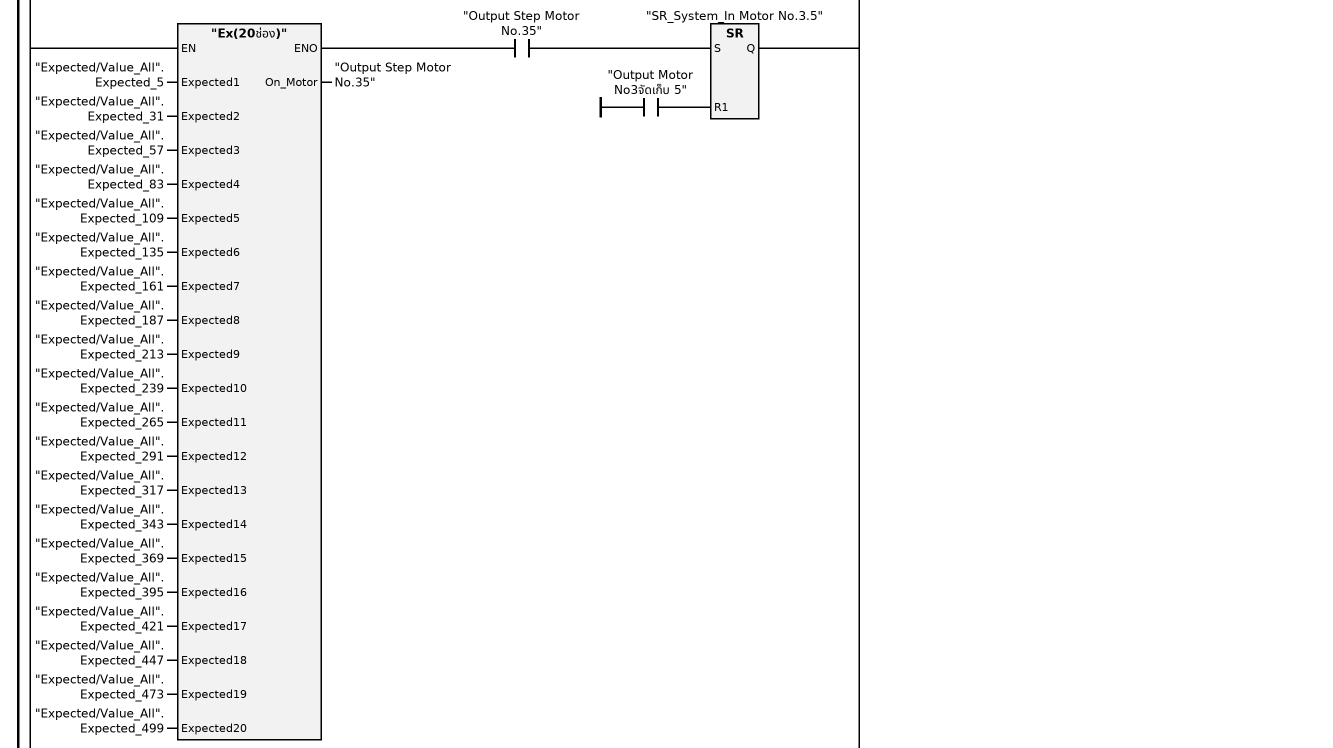
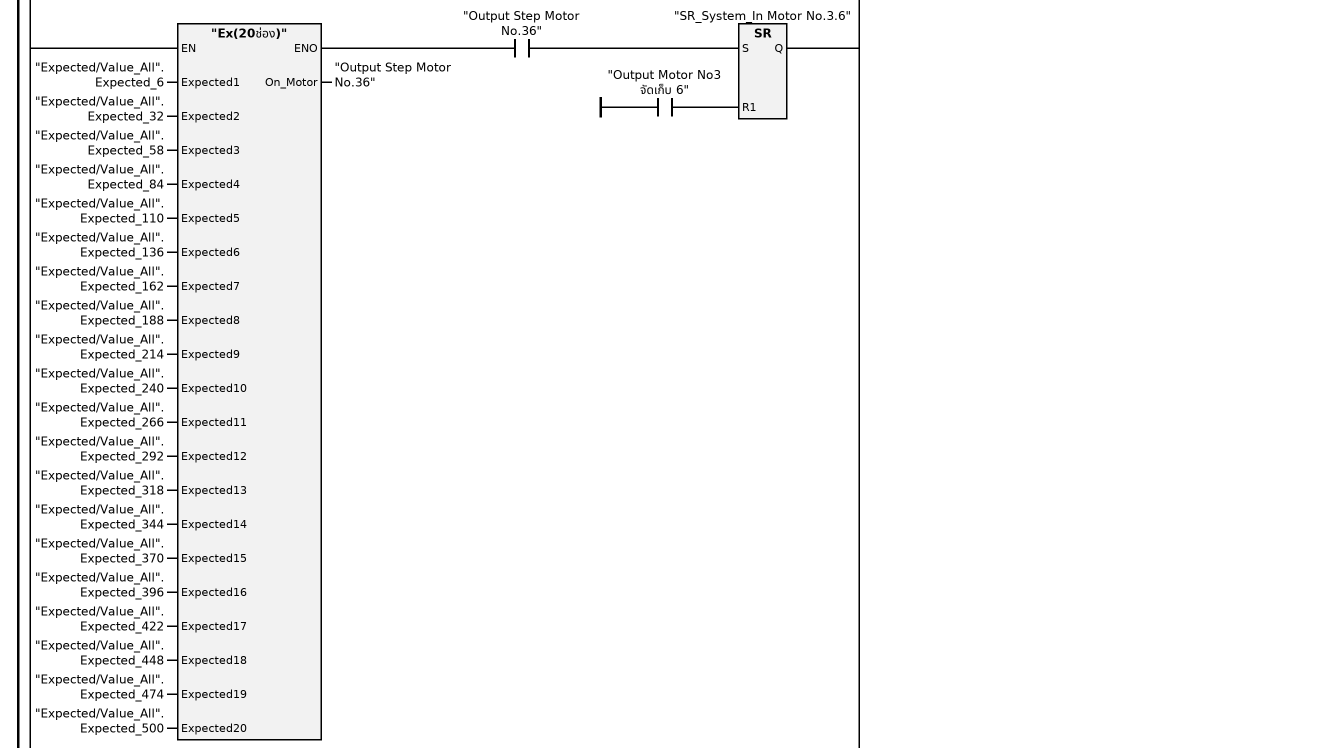
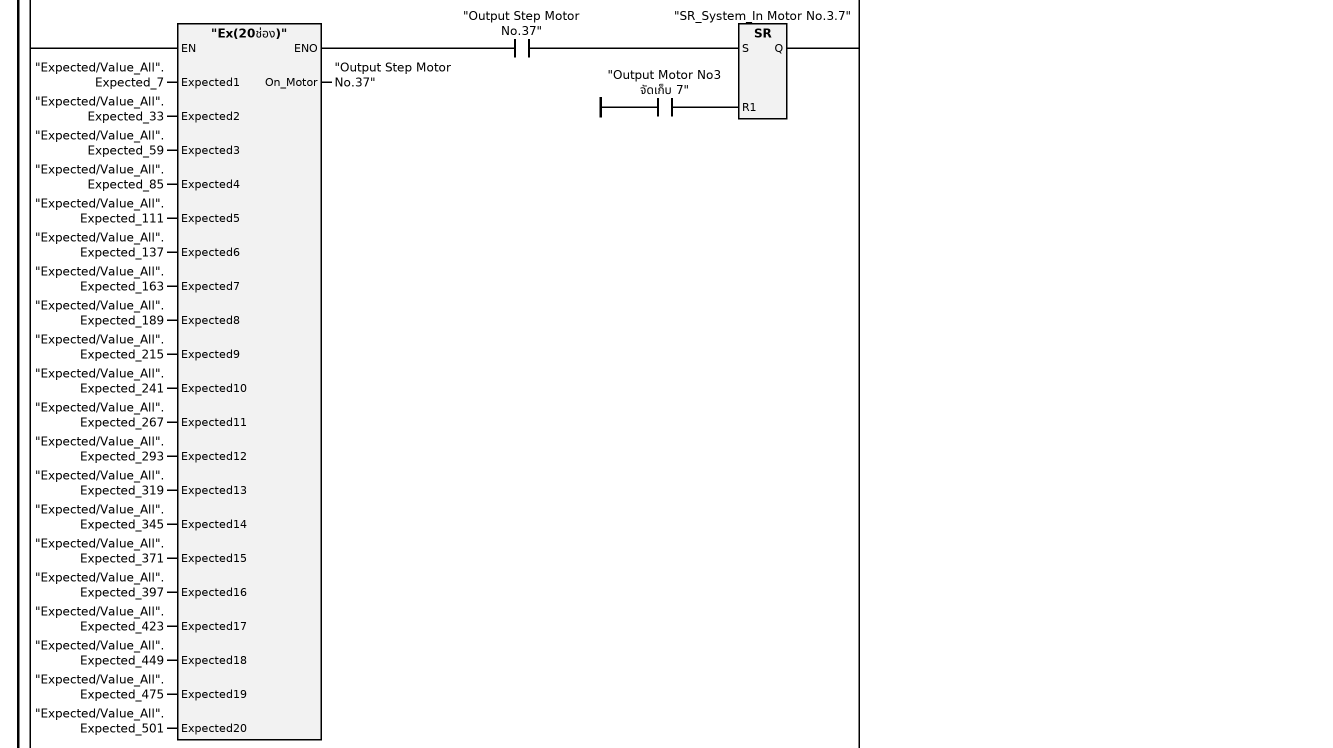
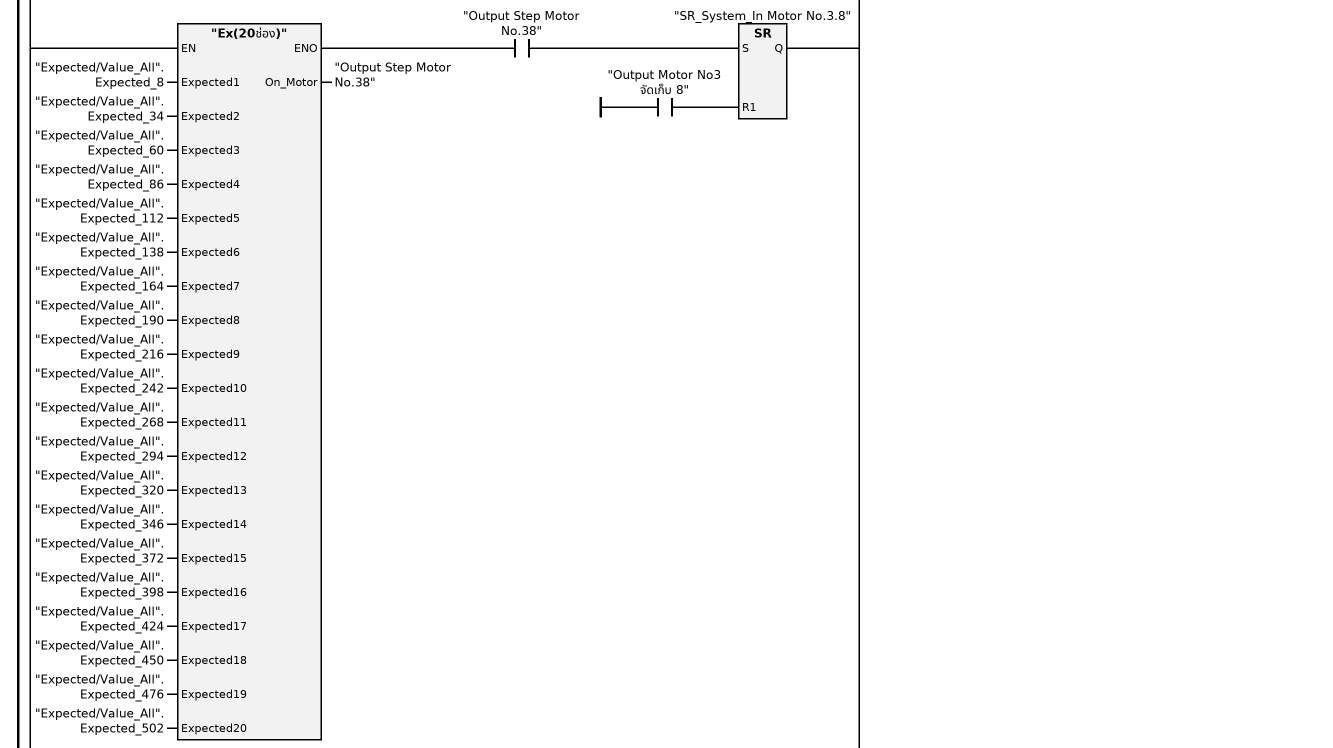
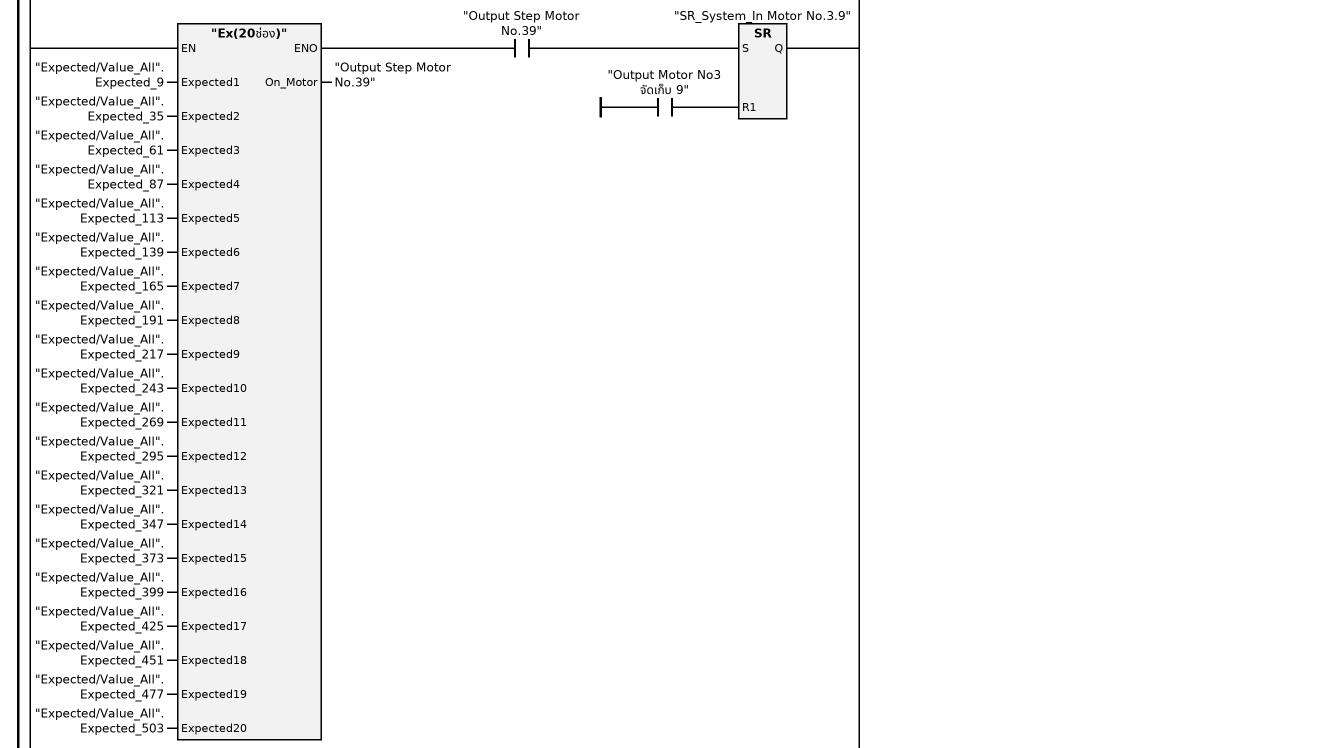
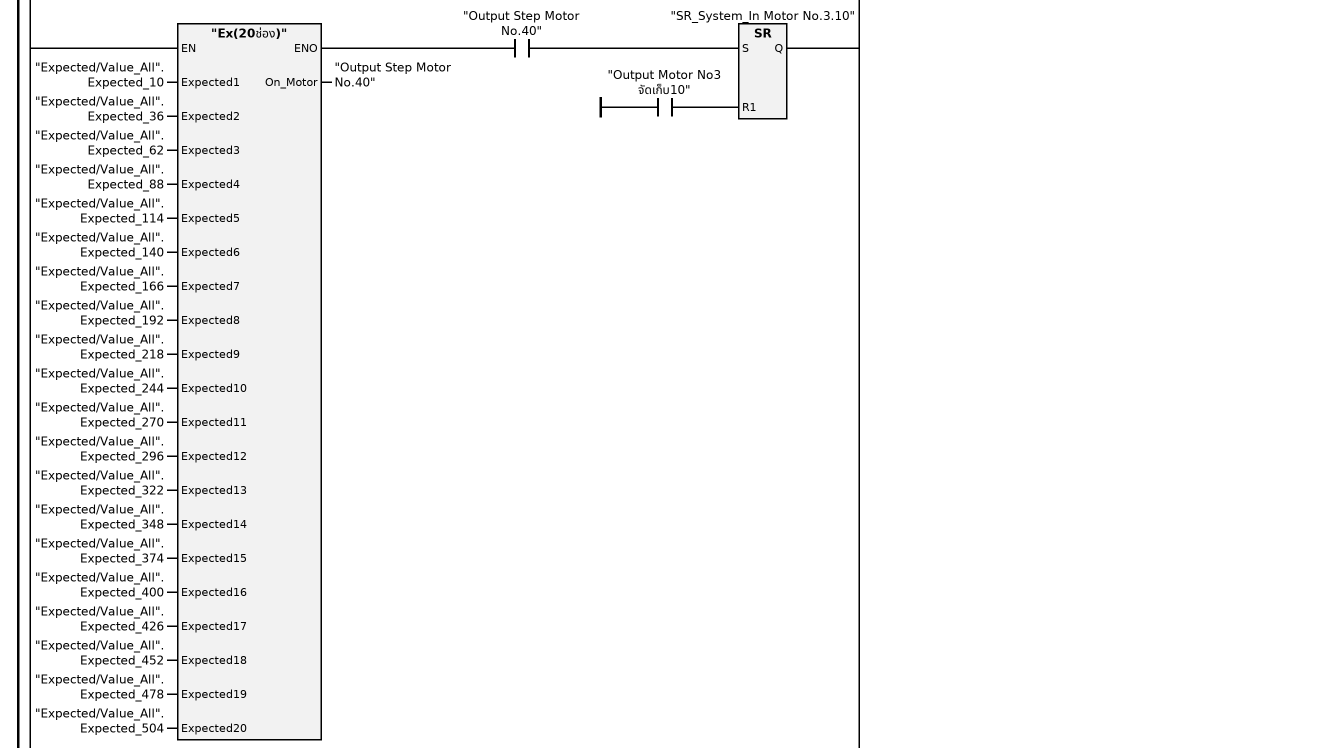
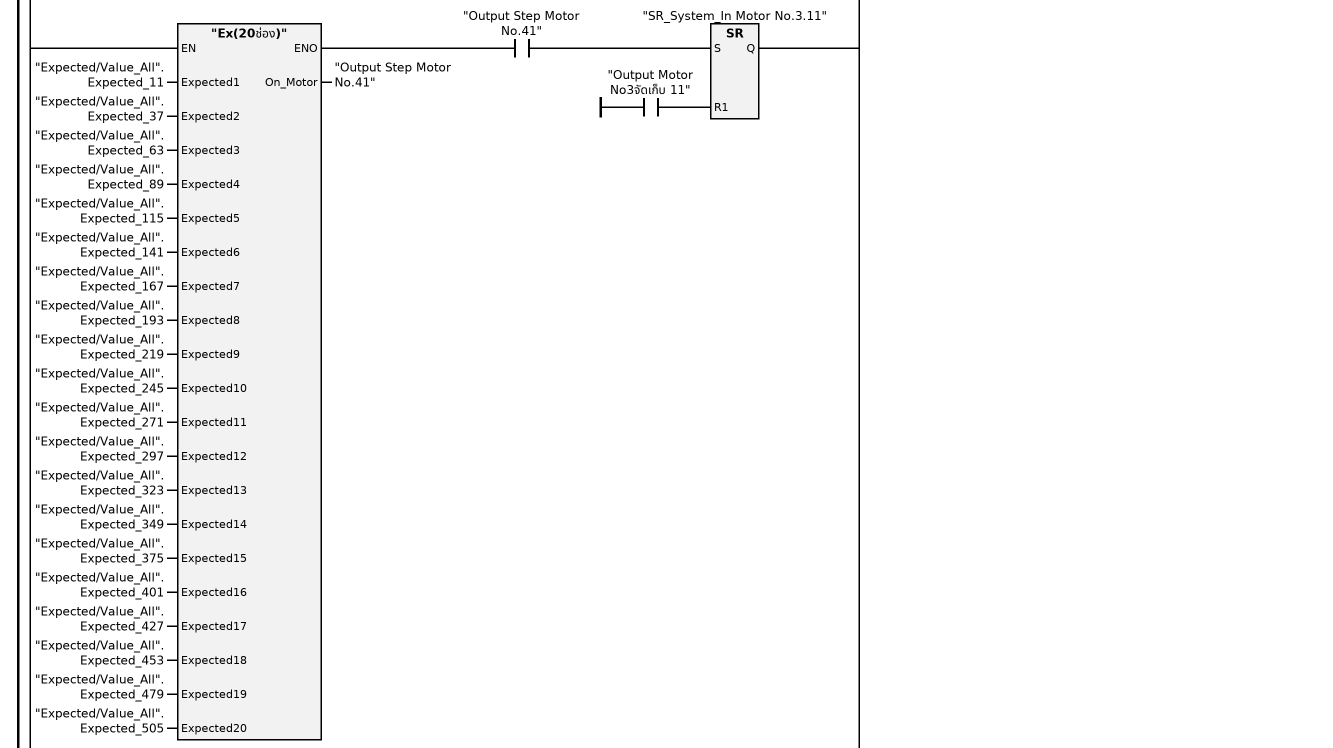
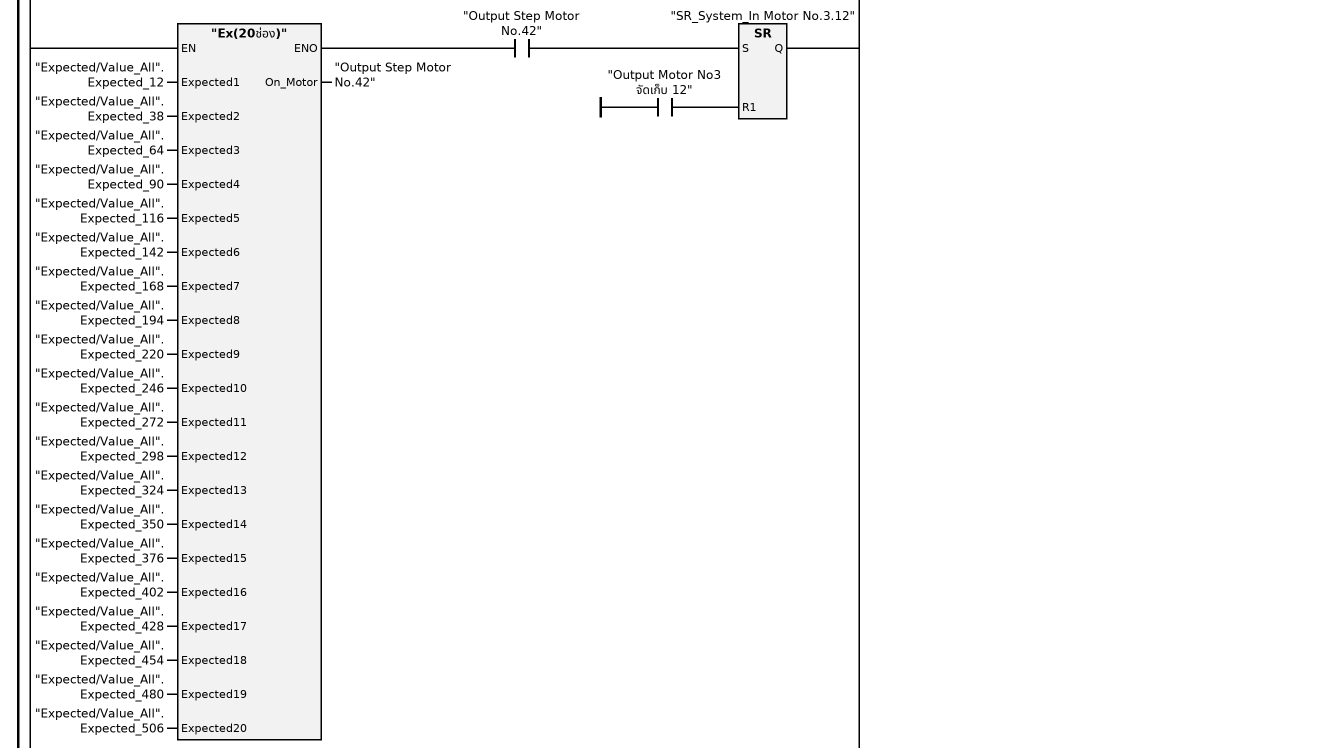
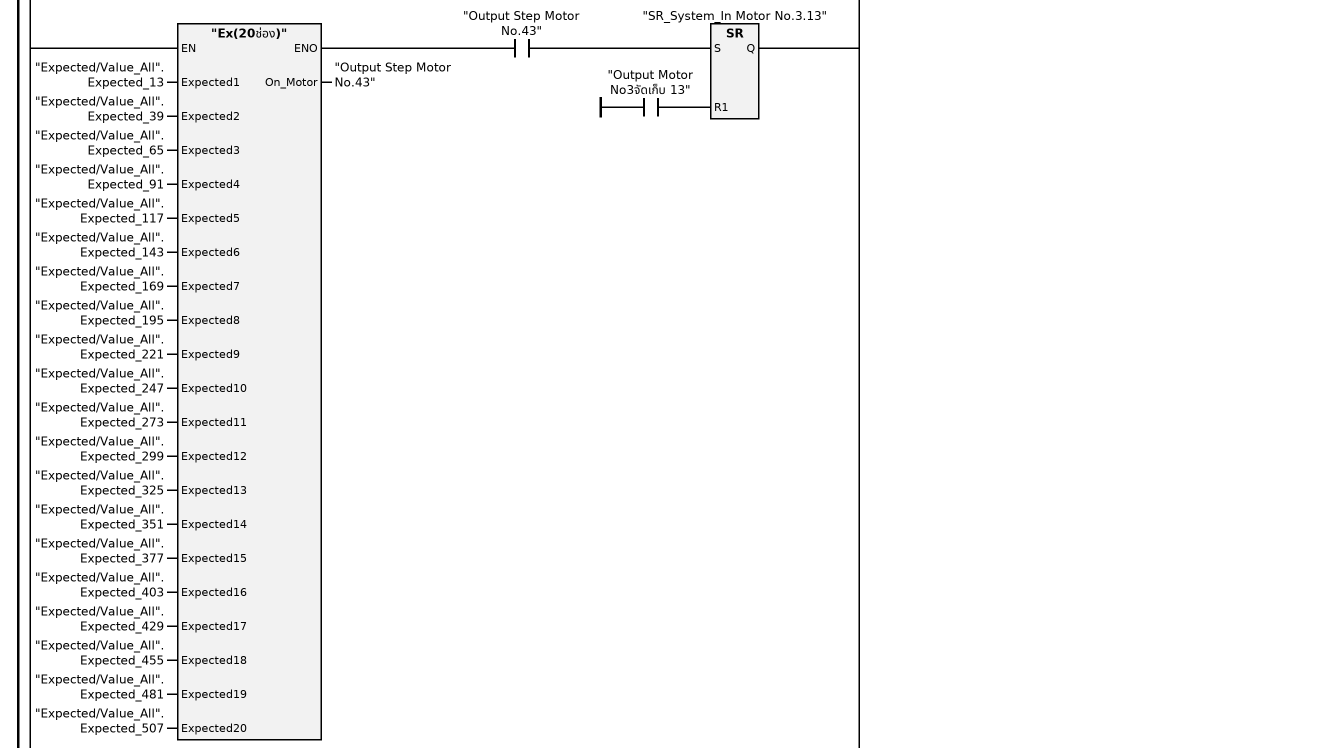
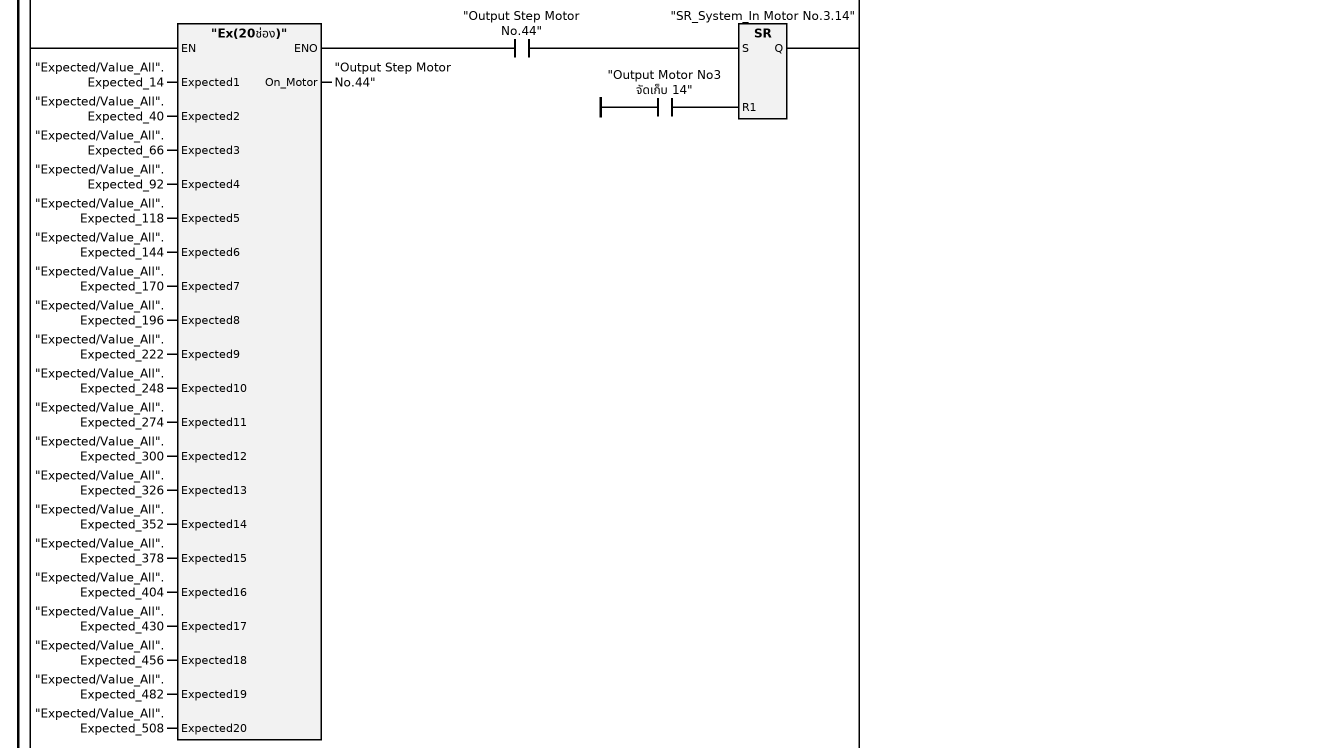
